Yaskawa INFORM job: THAPPY.JBI

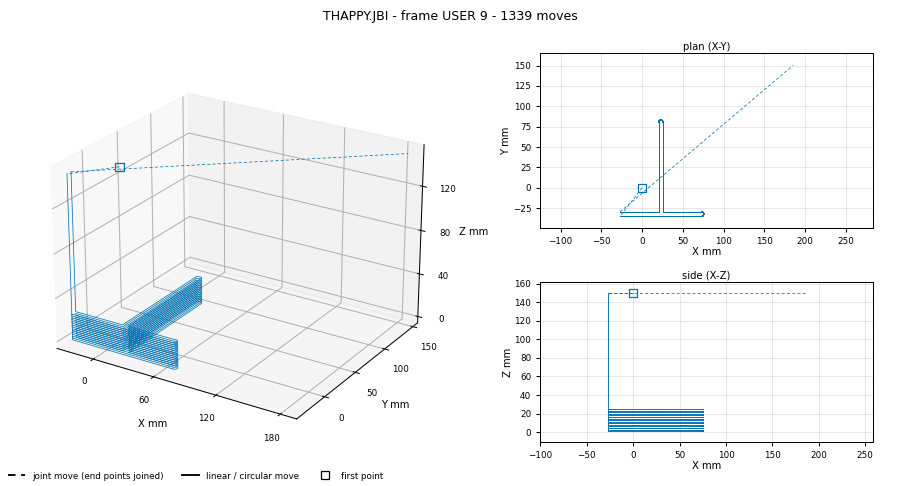
[picture p0: tool path of THAPPY.JBI in frame USER 9, 1339 of 1369 moves have a stored position in this frame; points joined in program order, loops and branches not executed]
/JOB
//NAME TTEST
//POS
///NPOS 1369,0,0,0,0,0
///USER 9
///TOOL 1
///POSTYPE USER
///RECTAN
///RCONF 1,0,0,0,0,0,0,0,0,0,0,0,0,0,0,0,0,0,0,0,0,0,0,0
C00000=0.000,0.000,150.000,0.0000,0.0000,-170.0000
C00001=-27.000,-35.000,150.000,0.0000,0.0000,-170.0000
C00002=-27.000,-35.000,1.000,0.0000,0.0000,-170.0000
C00003=-22.000,-35.000,1.000,0.0000,0.0000,-170.0000
C00004=-17.000,-35.000,1.000,0.0000,0.0000,-170.0000
C00005=-12.000,-35.000,1.000,0.0000,0.0000,-170.0000
C00006=-7.000,-35.000,1.000,0.0000,0.0000,-170.0000
C00007=-2.000,-35.000,1.000,0.0000,0.0000,-170.0000
C00008=3.000,-35.000,1.000,0.0000,0.0000,-170.0000
C00009=8.000,-35.000,1.000,0.0000,0.0000,-170.0000
C00010=13.000,-35.000,1.000,0.0000,0.0000,-170.0000
C00011=18.000,-35.000,1.000,0.0000,0.0000,-170.0000
C00012=23.000,-35.000,1.000,0.0000,0.0000,-170.0000
C00013=28.000,-35.000,1.000,0.0000,0.0000,-170.0000
C00014=33.000,-35.000,1.000,0.0000,0.0000,-170.0000
C00015=38.000,-35.000,1.000,0.0000,0.0000,-170.0000
C00016=43.000,-35.000,1.000,0.0000,0.0000,-170.0000
C00017=48.000,-35.000,1.000,0.0000,0.0000,-170.0000
C00018=53.000,-35.000,1.000,0.0000,0.0000,-170.0000
C00019=58.000,-35.000,1.000,0.0000,0.0000,-170.0000
C00020=63.000,-35.000,1.000,0.0000,0.0000,-170.0000
C00021=68.000,-35.000,1.000,0.0000,0.0000,-170.0000
C00022=73.000,-35.000,1.000,0.0000,0.0000,-170.0000
C00023=73.000,-35.000,1.000,0.0000,0.0000,-170.0000
C00024=75.750,-32.250,1.000,0.0000,0.0000,-170.0000
C00025=73.000,-29.500,1.000,0.0000,0.0000,-170.0000
C00026=68.275,-29.500,1.000,0.0000,0.0000,-170.0000
C00027=63.550,-29.500,1.000,0.0000,0.0000,-170.0000
C00028=58.825,-29.500,1.000,0.0000,0.0000,-170.0000
C00029=54.100,-29.500,1.000,0.0000,0.0000,-170.0000
C00030=49.375,-29.500,1.000,0.0000,0.0000,-170.0000
C00031=44.650,-29.500,1.000,0.0000,0.0000,-170.0000
C00032=39.925,-29.500,1.000,0.0000,0.0000,-170.0000
C00033=35.200,-29.500,1.000,0.0000,0.0000,-170.0000
C00034=30.475,-29.500,1.000,0.0000,0.0000,-170.0000
C00035=25.750,-29.500,1.000,0.0000,0.0000,-170.0000
C00036=25.750,-24.500,1.000,0.0000,0.0000,-170.0000
C00037=25.750,-19.500,1.000,0.0000,0.0000,-170.0000
C00038=25.750,-14.500,1.000,0.0000,0.0000,-170.0000
C00039=25.750,-9.500,1.000,0.0000,0.0000,-170.0000
C00040=25.750,-4.500,1.000,0.0000,0.0000,-170.0000
C00041=25.750,0.500,1.000,0.0000,0.0000,-170.0000
C00042=25.750,5.500,1.000,0.0000,0.0000,-170.0000
C00043=25.750,10.500,1.000,0.0000,0.0000,-170.0000
C00044=25.750,15.500,1.000,0.0000,0.0000,-170.0000
C00045=25.750,20.500,1.000,0.0000,0.0000,-170.0000
C00046=25.750,25.500,1.000,0.0000,0.0000,-170.0000
C00047=25.750,30.500,1.000,0.0000,0.0000,-170.0000
C00048=25.750,35.500,1.000,0.0000,0.0000,-170.0000
C00049=25.750,40.500,1.000,0.0000,0.0000,-170.0000
C00050=25.750,45.500,1.000,0.0000,0.0000,-170.0000
C00051=25.750,50.500,1.000,0.0000,0.0000,-170.0000
C00052=25.750,55.500,1.000,0.0000,0.0000,-170.0000
C00053=25.750,60.500,1.000,0.0000,0.0000,-170.0000
C00054=25.750,65.500,1.000,0.0000,0.0000,-170.0000
C00055=25.750,70.500,1.000,0.0000,0.0000,-170.0000
C00056=25.750,75.500,1.000,0.0000,0.0000,-170.0000
C00057=25.750,80.500,1.000,0.0000,0.0000,-170.0000
C00058=25.750,80.500,1.000,0.0000,0.0000,-170.0000
C00059=23.000,83.250,1.000,0.0000,0.0000,-170.0000
C00060=20.250,80.500,1.000,0.0000,0.0000,-170.0000
C00061=20.250,75.500,1.000,0.0000,0.0000,-170.0000
C00062=20.250,70.500,1.000,0.0000,0.0000,-170.0000
C00063=20.250,65.500,1.000,0.0000,0.0000,-170.0000
C00064=20.250,60.500,1.000,0.0000,0.0000,-170.0000
C00065=20.250,55.500,1.000,0.0000,0.0000,-170.0000
C00066=20.250,50.500,1.000,0.0000,0.0000,-170.0000
C00067=20.250,45.500,1.000,0.0000,0.0000,-170.0000
C00068=20.250,40.500,1.000,0.0000,0.0000,-170.0000
C00069=20.250,35.500,1.000,0.0000,0.0000,-170.0000
C00070=20.250,30.500,1.000,0.0000,0.0000,-170.0000
C00071=20.250,25.500,1.000,0.0000,0.0000,-170.0000
C00072=20.250,20.500,1.000,0.0000,0.0000,-170.0000
C00073=20.250,15.500,1.000,0.0000,0.0000,-170.0000
C00074=20.250,10.500,1.000,0.0000,0.0000,-170.0000
C00075=20.250,5.500,1.000,0.0000,0.0000,-170.0000
C00076=20.250,0.500,1.000,0.0000,0.0000,-170.0000
C00077=20.250,-4.500,1.000,0.0000,0.0000,-170.0000
C00078=20.250,-9.500,1.000,0.0000,0.0000,-170.0000
C00079=20.250,-14.500,1.000,0.0000,0.0000,-170.0000
C00080=20.250,-19.500,1.000,0.0000,0.0000,-170.0000
C00081=20.250,-24.500,1.000,0.0000,0.0000,-170.0000
C00082=20.250,-29.500,1.000,0.0000,0.0000,-170.0000
C00083=15.525,-29.500,1.000,0.0000,0.0000,-170.0000
C00084=10.800,-29.500,1.000,0.0000,0.0000,-170.0000
C00085=6.075,-29.500,1.000,0.0000,0.0000,-170.0000
C00086=1.350,-29.500,1.000,0.0000,0.0000,-170.0000
C00087=-3.375,-29.500,1.000,0.0000,0.0000,-170.0000
C00088=-8.100,-29.500,1.000,0.0000,0.0000,-170.0000
C00089=-12.825,-29.500,1.000,0.0000,0.0000,-170.0000
C00090=-17.550,-29.500,1.000,0.0000,0.0000,-170.0000
C00091=-22.275,-29.500,1.000,0.0000,0.0000,-170.0000
C00092=-27.000,-29.500,1.000,0.0000,0.0000,-170.0000
C00093=-27.000,-29.500,2.700,0.0000,0.0000,-170.0000
C00094=-22.275,-29.500,2.700,0.0000,0.0000,-170.0000
C00095=-17.550,-29.500,2.700,0.0000,0.0000,-170.0000
C00096=-12.825,-29.500,2.700,0.0000,0.0000,-170.0000
C00097=-8.100,-29.500,2.700,0.0000,0.0000,-170.0000
C00098=-3.375,-29.500,2.700,0.0000,0.0000,-170.0000
C00099=1.350,-29.500,2.700,0.0000,0.0000,-170.0000
C00100=6.075,-29.500,2.700,0.0000,0.0000,-170.0000
C00101=10.800,-29.500,2.700,0.0000,0.0000,-170.0000
C00102=15.525,-29.500,2.700,0.0000,0.0000,-170.0000
C00103=20.250,-29.500,2.700,0.0000,0.0000,-170.0000
C00104=20.250,-24.500,2.700,0.0000,0.0000,-170.0000
C00105=20.250,-19.500,2.700,0.0000,0.0000,-170.0000
C00106=20.250,-14.500,2.700,0.0000,0.0000,-170.0000
C00107=20.250,-9.500,2.700,0.0000,0.0000,-170.0000
C00108=20.250,-4.500,2.700,0.0000,0.0000,-170.0000
C00109=20.250,0.500,2.700,0.0000,0.0000,-170.0000
C00110=20.250,5.500,2.700,0.0000,0.0000,-170.0000
C00111=20.250,10.500,2.700,0.0000,0.0000,-170.0000
C00112=20.250,15.500,2.700,0.0000,0.0000,-170.0000
C00113=20.250,20.500,2.700,0.0000,0.0000,-170.0000
C00114=20.250,25.500,2.700,0.0000,0.0000,-170.0000
C00115=20.250,30.500,2.700,0.0000,0.0000,-170.0000
C00116=20.250,35.500,2.700,0.0000,0.0000,-170.0000
C00117=20.250,40.500,2.700,0.0000,0.0000,-170.0000
C00118=20.250,45.500,2.700,0.0000,0.0000,-170.0000
C00119=20.250,50.500,2.700,0.0000,0.0000,-170.0000
C00120=20.250,55.500,2.700,0.0000,0.0000,-170.0000
C00121=20.250,60.500,2.700,0.0000,0.0000,-170.0000
C00122=20.250,65.500,2.700,0.0000,0.0000,-170.0000
C00123=20.250,70.500,2.700,0.0000,0.0000,-170.0000
C00124=20.250,75.500,2.700,0.0000,0.0000,-170.0000
C00125=20.250,80.500,2.700,0.0000,0.0000,-170.0000
C00126=20.250,80.500,2.700,0.0000,0.0000,-170.0000
C00127=23.000,83.250,2.700,0.0000,0.0000,-170.0000
C00128=25.750,80.500,2.700,0.0000,0.0000,-170.0000
C00129=25.750,75.500,2.700,0.0000,0.0000,-170.0000
C00130=25.750,70.500,2.700,0.0000,0.0000,-170.0000
C00131=25.750,65.500,2.700,0.0000,0.0000,-170.0000
C00132=25.750,60.500,2.700,0.0000,0.0000,-170.0000
C00133=25.750,55.500,2.700,0.0000,0.0000,-170.0000
C00134=25.750,50.500,2.700,0.0000,0.0000,-170.0000
C00135=25.750,45.500,2.700,0.0000,0.0000,-170.0000
C00136=25.750,40.500,2.700,0.0000,0.0000,-170.0000
C00137=25.750,35.500,2.700,0.0000,0.0000,-170.0000
C00138=25.750,30.500,2.700,0.0000,0.0000,-170.0000
C00139=25.750,25.500,2.700,0.0000,0.0000,-170.0000
C00140=25.750,20.500,2.700,0.0000,0.0000,-170.0000
C00141=25.750,15.500,2.700,0.0000,0.0000,-170.0000
C00142=25.750,10.500,2.700,0.0000,0.0000,-170.0000
C00143=25.750,5.500,2.700,0.0000,0.0000,-170.0000
C00144=25.750,0.500,2.700,0.0000,0.0000,-170.0000
C00145=25.750,-4.500,2.700,0.0000,0.0000,-170.0000
C00146=25.750,-9.500,2.700,0.0000,0.0000,-170.0000
C00147=25.750,-14.500,2.700,0.0000,0.0000,-170.0000
C00148=25.750,-19.500,2.700,0.0000,0.0000,-170.0000
C00149=25.750,-24.500,2.700,0.0000,0.0000,-170.0000
C00150=25.750,-29.500,2.700,0.0000,0.0000,-170.0000
C00151=30.475,-29.500,2.700,0.0000,0.0000,-170.0000
C00152=35.200,-29.500,2.700,0.0000,0.0000,-170.0000
C00153=39.925,-29.500,2.700,0.0000,0.0000,-170.0000
C00154=44.650,-29.500,2.700,0.0000,0.0000,-170.0000
C00155=49.375,-29.500,2.700,0.0000,0.0000,-170.0000
C00156=54.100,-29.500,2.700,0.0000,0.0000,-170.0000
C00157=58.825,-29.500,2.700,0.0000,0.0000,-170.0000
C00158=63.550,-29.500,2.700,0.0000,0.0000,-170.0000
C00159=68.275,-29.500,2.700,0.0000,0.0000,-170.0000
C00160=73.000,-29.500,2.700,0.0000,0.0000,-170.0000
C00161=73.000,-29.500,2.700,0.0000,0.0000,-170.0000
C00162=75.750,-32.250,2.700,0.0000,0.0000,-170.0000
C00163=73.000,-35.000,2.700,0.0000,0.0000,-170.0000
C00164=68.000,-35.000,2.700,0.0000,0.0000,-170.0000
C00165=63.000,-35.000,2.700,0.0000,0.0000,-170.0000
C00166=58.000,-35.000,2.700,0.0000,0.0000,-170.0000
C00167=53.000,-35.000,2.700,0.0000,0.0000,-170.0000
C00168=48.000,-35.000,2.700,0.0000,0.0000,-170.0000
C00169=43.000,-35.000,2.700,0.0000,0.0000,-170.0000
C00170=38.000,-35.000,2.700,0.0000,0.0000,-170.0000
C00171=33.000,-35.000,2.700,0.0000,0.0000,-170.0000
C00172=28.000,-35.000,2.700,0.0000,0.0000,-170.0000
C00173=23.000,-35.000,2.700,0.0000,0.0000,-170.0000
C00174=18.000,-35.000,2.700,0.0000,0.0000,-170.0000
C00175=13.000,-35.000,2.700,0.0000,0.0000,-170.0000
C00176=8.000,-35.000,2.700,0.0000,0.0000,-170.0000
C00177=3.000,-35.000,2.700,0.0000,0.0000,-170.0000
C00178=-2.000,-35.000,2.700,0.0000,0.0000,-170.0000
C00179=-7.000,-35.000,2.700,0.0000,0.0000,-170.0000
C00180=-12.000,-35.000,2.700,0.0000,0.0000,-170.0000
C00181=-17.000,-35.000,2.700,0.0000,0.0000,-170.0000
C00182=-22.000,-35.000,2.700,0.0000,0.0000,-170.0000
C00183=-27.000,-35.000,2.700,0.0000,0.0000,-170.0000
C00184=-27.000,-35.000,4.400,0.0000,0.0000,-170.0000
C00185=-22.000,-35.000,4.400,0.0000,0.0000,-170.0000
C00186=-17.000,-35.000,4.400,0.0000,0.0000,-170.0000
C00187=-12.000,-35.000,4.400,0.0000,0.0000,-170.0000
C00188=-7.000,-35.000,4.400,0.0000,0.0000,-170.0000
C00189=-2.000,-35.000,4.400,0.0000,0.0000,-170.0000
C00190=3.000,-35.000,4.400,0.0000,0.0000,-170.0000
C00191=8.000,-35.000,4.400,0.0000,0.0000,-170.0000
C00192=13.000,-35.000,4.400,0.0000,0.0000,-170.0000
C00193=18.000,-35.000,4.400,0.0000,0.0000,-170.0000
C00194=23.000,-35.000,4.400,0.0000,0.0000,-170.0000
C00195=28.000,-35.000,4.400,0.0000,0.0000,-170.0000
C00196=33.000,-35.000,4.400,0.0000,0.0000,-170.0000
C00197=38.000,-35.000,4.400,0.0000,0.0000,-170.0000
C00198=43.000,-35.000,4.400,0.0000,0.0000,-170.0000
C00199=48.000,-35.000,4.400,0.0000,0.0000,-170.0000
C00200=53.000,-35.000,4.400,0.0000,0.0000,-170.0000
C00201=58.000,-35.000,4.400,0.0000,0.0000,-170.0000
C00202=63.000,-35.000,4.400,0.0000,0.0000,-170.0000
C00203=68.000,-35.000,4.400,0.0000,0.0000,-170.0000
C00204=73.000,-35.000,4.400,0.0000,0.0000,-170.0000
C00205=73.000,-35.000,4.400,0.0000,0.0000,-170.0000
C00206=75.750,-32.250,4.400,0.0000,0.0000,-170.0000
C00207=73.000,-29.500,4.400,0.0000,0.0000,-170.0000
C00208=68.275,-29.500,4.400,0.0000,0.0000,-170.0000
C00209=63.550,-29.500,4.400,0.0000,0.0000,-170.0000
C00210=58.825,-29.500,4.400,0.0000,0.0000,-170.0000
C00211=54.100,-29.500,4.400,0.0000,0.0000,-170.0000
C00212=49.375,-29.500,4.400,0.0000,0.0000,-170.0000
C00213=44.650,-29.500,4.400,0.0000,0.0000,-170.0000
C00214=39.925,-29.500,4.400,0.0000,0.0000,-170.0000
C00215=35.200,-29.500,4.400,0.0000,0.0000,-170.0000
C00216=30.475,-29.500,4.400,0.0000,0.0000,-170.0000
C00217=25.750,-29.500,4.400,0.0000,0.0000,-170.0000
C00218=25.750,-24.500,4.400,0.0000,0.0000,-170.0000
C00219=25.750,-19.500,4.400,0.0000,0.0000,-170.0000
C00220=25.750,-14.500,4.400,0.0000,0.0000,-170.0000
C00221=25.750,-9.500,4.400,0.0000,0.0000,-170.0000
C00222=25.750,-4.500,4.400,0.0000,0.0000,-170.0000
C00223=25.750,0.500,4.400,0.0000,0.0000,-170.0000
C00224=25.750,5.500,4.400,0.0000,0.0000,-170.0000
C00225=25.750,10.500,4.400,0.0000,0.0000,-170.0000
C00226=25.750,15.500,4.400,0.0000,0.0000,-170.0000
C00227=25.750,20.500,4.400,0.0000,0.0000,-170.0000
C00228=25.750,25.500,4.400,0.0000,0.0000,-170.0000
C00229=25.750,30.500,4.400,0.0000,0.0000,-170.0000
C00230=25.750,35.500,4.400,0.0000,0.0000,-170.0000
C00231=25.750,40.500,4.400,0.0000,0.0000,-170.0000
C00232=25.750,45.500,4.400,0.0000,0.0000,-170.0000
C00233=25.750,50.500,4.400,0.0000,0.0000,-170.0000
C00234=25.750,55.500,4.400,0.0000,0.0000,-170.0000
C00235=25.750,60.500,4.400,0.0000,0.0000,-170.0000
C00236=25.750,65.500,4.400,0.0000,0.0000,-170.0000
C00237=25.750,70.500,4.400,0.0000,0.0000,-170.0000
C00238=25.750,75.500,4.400,0.0000,0.0000,-170.0000
C00239=25.750,80.500,4.400,0.0000,0.0000,-170.0000
C00240=25.750,80.500,4.400,0.0000,0.0000,-170.0000
C00241=23.000,83.250,4.400,0.0000,0.0000,-170.0000
C00242=20.250,80.500,4.400,0.0000,0.0000,-170.0000
C00243=20.250,75.500,4.400,0.0000,0.0000,-170.0000
C00244=20.250,70.500,4.400,0.0000,0.0000,-170.0000
C00245=20.250,65.500,4.400,0.0000,0.0000,-170.0000
C00246=20.250,60.500,4.400,0.0000,0.0000,-170.0000
C00247=20.250,55.500,4.400,0.0000,0.0000,-170.0000
C00248=20.250,50.500,4.400,0.0000,0.0000,-170.0000
C00249=20.250,45.500,4.400,0.0000,0.0000,-170.0000
C00250=20.250,40.500,4.400,0.0000,0.0000,-170.0000
C00251=20.250,35.500,4.400,0.0000,0.0000,-170.0000
C00252=20.250,30.500,4.400,0.0000,0.0000,-170.0000
C00253=20.250,25.500,4.400,0.0000,0.0000,-170.0000
C00254=20.250,20.500,4.400,0.0000,0.0000,-170.0000
C00255=20.250,15.500,4.400,0.0000,0.0000,-170.0000
C00256=20.250,10.500,4.400,0.0000,0.0000,-170.0000
C00257=20.250,5.500,4.400,0.0000,0.0000,-170.0000
C00258=20.250,0.500,4.400,0.0000,0.0000,-170.0000
C00259=20.250,-4.500,4.400,0.0000,0.0000,-170.0000
C00260=20.250,-9.500,4.400,0.0000,0.0000,-170.0000
C00261=20.250,-14.500,4.400,0.0000,0.0000,-170.0000
C00262=20.250,-19.500,4.400,0.0000,0.0000,-170.0000
C00263=20.250,-24.500,4.400,0.0000,0.0000,-170.0000
C00264=20.250,-29.500,4.400,0.0000,0.0000,-170.0000
C00265=15.525,-29.500,4.400,0.0000,0.0000,-170.0000
C00266=10.800,-29.500,4.400,0.0000,0.0000,-170.0000
C00267=6.075,-29.500,4.400,0.0000,0.0000,-170.0000
C00268=1.350,-29.500,4.400,0.0000,0.0000,-170.0000
C00269=-3.375,-29.500,4.400,0.0000,0.0000,-170.0000
C00270=-8.100,-29.500,4.400,0.0000,0.0000,-170.0000
C00271=-12.825,-29.500,4.400,0.0000,0.0000,-170.0000
C00272=-17.550,-29.500,4.400,0.0000,0.0000,-170.0000
C00273=-22.275,-29.500,4.400,0.0000,0.0000,-170.0000
C00274=-27.000,-29.500,4.400,0.0000,0.0000,-170.0000
C00275=-27.000,-29.500,6.100,0.0000,0.0000,-170.0000
C00276=-22.275,-29.500,6.100,0.0000,0.0000,-170.0000
C00277=-17.550,-29.500,6.100,0.0000,0.0000,-170.0000
C00278=-12.825,-29.500,6.100,0.0000,0.0000,-170.0000
C00279=-8.100,-29.500,6.100,0.0000,0.0000,-170.0000
C00280=-3.375,-29.500,6.100,0.0000,0.0000,-170.0000
C00281=1.350,-29.500,6.100,0.0000,0.0000,-170.0000
C00282=6.075,-29.500,6.100,0.0000,0.0000,-170.0000
C00283=10.800,-29.500,6.100,0.0000,0.0000,-170.0000
C00284=15.525,-29.500,6.100,0.0000,0.0000,-170.0000
C00285=20.250,-29.500,6.100,0.0000,0.0000,-170.0000
C00286=20.250,-24.500,6.100,0.0000,0.0000,-170.0000
C00287=20.250,-19.500,6.100,0.0000,0.0000,-170.0000
C00288=20.250,-14.500,6.100,0.0000,0.0000,-170.0000
C00289=20.250,-9.500,6.100,0.0000,0.0000,-170.0000
C00290=20.250,-4.500,6.100,0.0000,0.0000,-170.0000
C00291=20.250,0.500,6.100,0.0000,0.0000,-170.0000
C00292=20.250,5.500,6.100,0.0000,0.0000,-170.0000
C00293=20.250,10.500,6.100,0.0000,0.0000,-170.0000
C00294=20.250,15.500,6.100,0.0000,0.0000,-170.0000
C00295=20.250,20.500,6.100,0.0000,0.0000,-170.0000
C00296=20.250,25.500,6.100,0.0000,0.0000,-170.0000
C00297=20.250,30.500,6.100,0.0000,0.0000,-170.0000
C00298=20.250,35.500,6.100,0.0000,0.0000,-170.0000
C00299=20.250,40.500,6.100,0.0000,0.0000,-170.0000
C00300=20.250,45.500,6.100,0.0000,0.0000,-170.0000
C00301=20.250,50.500,6.100,0.0000,0.0000,-170.0000
C00302=20.250,55.500,6.100,0.0000,0.0000,-170.0000
C00303=20.250,60.500,6.100,0.0000,0.0000,-170.0000
C00304=20.250,65.500,6.100,0.0000,0.0000,-170.0000
C00305=20.250,70.500,6.100,0.0000,0.0000,-170.0000
C00306=20.250,75.500,6.100,0.0000,0.0000,-170.0000
C00307=20.250,80.500,6.100,0.0000,0.0000,-170.0000
C00308=20.250,80.500,6.100,0.0000,0.0000,-170.0000
C00309=23.000,83.250,6.100,0.0000,0.0000,-170.0000
C00310=25.750,80.500,6.100,0.0000,0.0000,-170.0000
C00311=25.750,75.500,6.100,0.0000,0.0000,-170.0000
C00312=25.750,70.500,6.100,0.0000,0.0000,-170.0000
C00313=25.750,65.500,6.100,0.0000,0.0000,-170.0000
C00314=25.750,60.500,6.100,0.0000,0.0000,-170.0000
C00315=25.750,55.500,6.100,0.0000,0.0000,-170.0000
C00316=25.750,50.500,6.100,0.0000,0.0000,-170.0000
C00317=25.750,45.500,6.100,0.0000,0.0000,-170.0000
C00318=25.750,40.500,6.100,0.0000,0.0000,-170.0000
C00319=25.750,35.500,6.100,0.0000,0.0000,-170.0000
C00320=25.750,30.500,6.100,0.0000,0.0000,-170.0000
C00321=25.750,25.500,6.100,0.0000,0.0000,-170.0000
C00322=25.750,20.500,6.100,0.0000,0.0000,-170.0000
C00323=25.750,15.500,6.100,0.0000,0.0000,-170.0000
C00324=25.750,10.500,6.100,0.0000,0.0000,-170.0000
C00325=25.750,5.500,6.100,0.0000,0.0000,-170.0000
C00326=25.750,0.500,6.100,0.0000,0.0000,-170.0000
C00327=25.750,-4.500,6.100,0.0000,0.0000,-170.0000
C00328=25.750,-9.500,6.100,0.0000,0.0000,-170.0000
C00329=25.750,-14.500,6.100,0.0000,0.0000,-170.0000
C00330=25.750,-19.500,6.100,0.0000,0.0000,-170.0000
C00331=25.750,-24.500,6.100,0.0000,0.0000,-170.0000
C00332=25.750,-29.500,6.100,0.0000,0.0000,-170.0000
C00333=30.475,-29.500,6.100,0.0000,0.0000,-170.0000
C00334=35.200,-29.500,6.100,0.0000,0.0000,-170.0000
C00335=39.925,-29.500,6.100,0.0000,0.0000,-170.0000
C00336=44.650,-29.500,6.100,0.0000,0.0000,-170.0000
C00337=49.375,-29.500,6.100,0.0000,0.0000,-170.0000
C00338=54.100,-29.500,6.100,0.0000,0.0000,-170.0000
C00339=58.825,-29.500,6.100,0.0000,0.0000,-170.0000
C00340=63.550,-29.500,6.100,0.0000,0.0000,-170.0000
C00341=68.275,-29.500,6.100,0.0000,0.0000,-170.0000
C00342=73.000,-29.500,6.100,0.0000,0.0000,-170.0000
C00343=73.000,-29.500,6.100,0.0000,0.0000,-170.0000
C00344=75.750,-32.250,6.100,0.0000,0.0000,-170.0000
C00345=73.000,-35.000,6.100,0.0000,0.0000,-170.0000
C00346=68.000,-35.000,6.100,0.0000,0.0000,-170.0000
C00347=63.000,-35.000,6.100,0.0000,0.0000,-170.0000
C00348=58.000,-35.000,6.100,0.0000,0.0000,-170.0000
C00349=53.000,-35.000,6.100,0.0000,0.0000,-170.0000
C00350=48.000,-35.000,6.100,0.0000,0.0000,-170.0000
C00351=43.000,-35.000,6.100,0.0000,0.0000,-170.0000
C00352=38.000,-35.000,6.100,0.0000,0.0000,-170.0000
C00353=33.000,-35.000,6.100,0.0000,0.0000,-170.0000
C00354=28.000,-35.000,6.100,0.0000,0.0000,-170.0000
C00355=23.000,-35.000,6.100,0.0000,0.0000,-170.0000
C00356=18.000,-35.000,6.100,0.0000,0.0000,-170.0000
C00357=13.000,-35.000,6.100,0.0000,0.0000,-170.0000
C00358=8.000,-35.000,6.100,0.0000,0.0000,-170.0000
C00359=3.000,-35.000,6.100,0.0000,0.0000,-170.0000
C00360=-2.000,-35.000,6.100,0.0000,0.0000,-170.0000
C00361=-7.000,-35.000,6.100,0.0000,0.0000,-170.0000
C00362=-12.000,-35.000,6.100,0.0000,0.0000,-170.0000
C00363=-17.000,-35.000,6.100,0.0000,0.0000,-170.0000
C00364=-22.000,-35.000,6.100,0.0000,0.0000,-170.0000
C00365=-27.000,-35.000,6.100,0.0000,0.0000,-170.0000
C00366=-27.000,-35.000,7.800,0.0000,0.0000,-170.0000
C00367=-22.000,-35.000,7.800,0.0000,0.0000,-170.0000
C00368=-17.000,-35.000,7.800,0.0000,0.0000,-170.0000
C00369=-12.000,-35.000,7.800,0.0000,0.0000,-170.0000
C00370=-7.000,-35.000,7.800,0.0000,0.0000,-170.0000
C00371=-2.000,-35.000,7.800,0.0000,0.0000,-170.0000
C00372=3.000,-35.000,7.800,0.0000,0.0000,-170.0000
C00373=8.000,-35.000,7.800,0.0000,0.0000,-170.0000
C00374=13.000,-35.000,7.800,0.0000,0.0000,-170.0000
C00375=18.000,-35.000,7.800,0.0000,0.0000,-170.0000
C00376=23.000,-35.000,7.800,0.0000,0.0000,-170.0000
C00377=28.000,-35.000,7.800,0.0000,0.0000,-170.0000
C00378=33.000,-35.000,7.800,0.0000,0.0000,-170.0000
C00379=38.000,-35.000,7.800,0.0000,0.0000,-170.0000
C00380=43.000,-35.000,7.800,0.0000,0.0000,-170.0000
C00381=48.000,-35.000,7.800,0.0000,0.0000,-170.0000
C00382=53.000,-35.000,7.800,0.0000,0.0000,-170.0000
C00383=58.000,-35.000,7.800,0.0000,0.0000,-170.0000
C00384=63.000,-35.000,7.800,0.0000,0.0000,-170.0000
C00385=68.000,-35.000,7.800,0.0000,0.0000,-170.0000
C00386=73.000,-35.000,7.800,0.0000,0.0000,-170.0000
C00387=73.000,-35.000,7.800,0.0000,0.0000,-170.0000
C00388=75.750,-32.250,7.800,0.0000,0.0000,-170.0000
C00389=73.000,-29.500,7.800,0.0000,0.0000,-170.0000
C00390=68.275,-29.500,7.800,0.0000,0.0000,-170.0000
C00391=63.550,-29.500,7.800,0.0000,0.0000,-170.0000
C00392=58.825,-29.500,7.800,0.0000,0.0000,-170.0000
C00393=54.100,-29.500,7.800,0.0000,0.0000,-170.0000
C00394=49.375,-29.500,7.800,0.0000,0.0000,-170.0000
C00395=44.650,-29.500,7.800,0.0000,0.0000,-170.0000
C00396=39.925,-29.500,7.800,0.0000,0.0000,-170.0000
C00397=35.200,-29.500,7.800,0.0000,0.0000,-170.0000
C00398=30.475,-29.500,7.800,0.0000,0.0000,-170.0000
C00399=25.750,-29.500,7.800,0.0000,0.0000,-170.0000
C00400=25.750,-24.500,7.800,0.0000,0.0000,-170.0000
C00401=25.750,-19.500,7.800,0.0000,0.0000,-170.0000
C00402=25.750,-14.500,7.800,0.0000,0.0000,-170.0000
C00403=25.750,-9.500,7.800,0.0000,0.0000,-170.0000
C00404=25.750,-4.500,7.800,0.0000,0.0000,-170.0000
C00405=25.750,0.500,7.800,0.0000,0.0000,-170.0000
C00406=25.750,5.500,7.800,0.0000,0.0000,-170.0000
C00407=25.750,10.500,7.800,0.0000,0.0000,-170.0000
C00408=25.750,15.500,7.800,0.0000,0.0000,-170.0000
C00409=25.750,20.500,7.800,0.0000,0.0000,-170.0000
C00410=25.750,25.500,7.800,0.0000,0.0000,-170.0000
C00411=25.750,30.500,7.800,0.0000,0.0000,-170.0000
C00412=25.750,35.500,7.800,0.0000,0.0000,-170.0000
C00413=25.750,40.500,7.800,0.0000,0.0000,-170.0000
C00414=25.750,45.500,7.800,0.0000,0.0000,-170.0000
C00415=25.750,50.500,7.800,0.0000,0.0000,-170.0000
C00416=25.750,55.500,7.800,0.0000,0.0000,-170.0000
C00417=25.750,60.500,7.800,0.0000,0.0000,-170.0000
C00418=25.750,65.500,7.800,0.0000,0.0000,-170.0000
C00419=25.750,70.500,7.800,0.0000,0.0000,-170.0000
C00420=25.750,75.500,7.800,0.0000,0.0000,-170.0000
C00421=25.750,80.500,7.800,0.0000,0.0000,-170.0000
C00422=25.750,80.500,7.800,0.0000,0.0000,-170.0000
C00423=23.000,83.250,7.800,0.0000,0.0000,-170.0000
C00424=20.250,80.500,7.800,0.0000,0.0000,-170.0000
C00425=20.250,75.500,7.800,0.0000,0.0000,-170.0000
C00426=20.250,70.500,7.800,0.0000,0.0000,-170.0000
C00427=20.250,65.500,7.800,0.0000,0.0000,-170.0000
C00428=20.250,60.500,7.800,0.0000,0.0000,-170.0000
C00429=20.250,55.500,7.800,0.0000,0.0000,-170.0000
C00430=20.250,50.500,7.800,0.0000,0.0000,-170.0000
C00431=20.250,45.500,7.800,0.0000,0.0000,-170.0000
C00432=20.250,40.500,7.800,0.0000,0.0000,-170.0000
C00433=20.250,35.500,7.800,0.0000,0.0000,-170.0000
C00434=20.250,30.500,7.800,0.0000,0.0000,-170.0000
C00435=20.250,25.500,7.800,0.0000,0.0000,-170.0000
C00436=20.250,20.500,7.800,0.0000,0.0000,-170.0000
C00437=20.250,15.500,7.800,0.0000,0.0000,-170.0000
C00438=20.250,10.500,7.800,0.0000,0.0000,-170.0000
C00439=20.250,5.500,7.800,0.0000,0.0000,-170.0000
C00440=20.250,0.500,7.800,0.0000,0.0000,-170.0000
C00441=20.250,-4.500,7.800,0.0000,0.0000,-170.0000
C00442=20.250,-9.500,7.800,0.0000,0.0000,-170.0000
C00443=20.250,-14.500,7.800,0.0000,0.0000,-170.0000
C00444=20.250,-19.500,7.800,0.0000,0.0000,-170.0000
C00445=20.250,-24.500,7.800,0.0000,0.0000,-170.0000
C00446=20.250,-29.500,7.800,0.0000,0.0000,-170.0000
C00447=15.525,-29.500,7.800,0.0000,0.0000,-170.0000
C00448=10.800,-29.500,7.800,0.0000,0.0000,-170.0000
C00449=6.075,-29.500,7.800,0.0000,0.0000,-170.0000
C00450=1.350,-29.500,7.800,0.0000,0.0000,-170.0000
C00451=-3.375,-29.500,7.800,0.0000,0.0000,-170.0000
C00452=-8.100,-29.500,7.800,0.0000,0.0000,-170.0000
C00453=-12.825,-29.500,7.800,0.0000,0.0000,-170.0000
C00454=-17.550,-29.500,7.800,0.0000,0.0000,-170.0000
C00455=-22.275,-29.500,7.800,0.0000,0.0000,-170.0000
C00456=-27.000,-29.500,7.800,0.0000,0.0000,-170.0000
C00457=-27.000,-29.500,9.500,0.0000,0.0000,-170.0000
C00458=-22.275,-29.500,9.500,0.0000,0.0000,-170.0000
C00459=-17.550,-29.500,9.500,0.0000,0.0000,-170.0000
C00460=-12.825,-29.500,9.500,0.0000,0.0000,-170.0000
C00461=-8.100,-29.500,9.500,0.0000,0.0000,-170.0000
C00462=-3.375,-29.500,9.500,0.0000,0.0000,-170.0000
C00463=1.350,-29.500,9.500,0.0000,0.0000,-170.0000
C00464=6.075,-29.500,9.500,0.0000,0.0000,-170.0000
C00465=10.800,-29.500,9.500,0.0000,0.0000,-170.0000
C00466=15.525,-29.500,9.500,0.0000,0.0000,-170.0000
C00467=20.250,-29.500,9.500,0.0000,0.0000,-170.0000
C00468=20.250,-24.500,9.500,0.0000,0.0000,-170.0000
C00469=20.250,-19.500,9.500,0.0000,0.0000,-170.0000
C00470=20.250,-14.500,9.500,0.0000,0.0000,-170.0000
C00471=20.250,-9.500,9.500,0.0000,0.0000,-170.0000
C00472=20.250,-4.500,9.500,0.0000,0.0000,-170.0000
C00473=20.250,0.500,9.500,0.0000,0.0000,-170.0000
C00474=20.250,5.500,9.500,0.0000,0.0000,-170.0000
C00475=20.250,10.500,9.500,0.0000,0.0000,-170.0000
C00476=20.250,15.500,9.500,0.0000,0.0000,-170.0000
C00477=20.250,20.500,9.500,0.0000,0.0000,-170.0000
C00478=20.250,25.500,9.500,0.0000,0.0000,-170.0000
C00479=20.250,30.500,9.500,0.0000,0.0000,-170.0000
C00480=20.250,35.500,9.500,0.0000,0.0000,-170.0000
C00481=20.250,40.500,9.500,0.0000,0.0000,-170.0000
C00482=20.250,45.500,9.500,0.0000,0.0000,-170.0000
C00483=20.250,50.500,9.500,0.0000,0.0000,-170.0000
C00484=20.250,55.500,9.500,0.0000,0.0000,-170.0000
C00485=20.250,60.500,9.500,0.0000,0.0000,-170.0000
C00486=20.250,65.500,9.500,0.0000,0.0000,-170.0000
C00487=20.250,70.500,9.500,0.0000,0.0000,-170.0000
C00488=20.250,75.500,9.500,0.0000,0.0000,-170.0000
C00489=20.250,80.500,9.500,0.0000,0.0000,-170.0000
C00490=20.250,80.500,9.500,0.0000,0.0000,-170.0000
C00491=23.000,83.250,9.500,0.0000,0.0000,-170.0000
C00492=25.750,80.500,9.500,0.0000,0.0000,-170.0000
C00493=25.750,75.500,9.500,0.0000,0.0000,-170.0000
C00494=25.750,70.500,9.500,0.0000,0.0000,-170.0000
C00495=25.750,65.500,9.500,0.0000,0.0000,-170.0000
C00496=25.750,60.500,9.500,0.0000,0.0000,-170.0000
C00497=25.750,55.500,9.500,0.0000,0.0000,-170.0000
C00498=25.750,50.500,9.500,0.0000,0.0000,-170.0000
C00499=25.750,45.500,9.500,0.0000,0.0000,-170.0000
C00500=25.750,40.500,9.500,0.0000,0.0000,-170.0000
C00501=25.750,35.500,9.500,0.0000,0.0000,-170.0000
C00502=25.750,30.500,9.500,0.0000,0.0000,-170.0000
C00503=25.750,25.500,9.500,0.0000,0.0000,-170.0000
C00504=25.750,20.500,9.500,0.0000,0.0000,-170.0000
C00505=25.750,15.500,9.500,0.0000,0.0000,-170.0000
C00506=25.750,10.500,9.500,0.0000,0.0000,-170.0000
C00507=25.750,5.500,9.500,0.0000,0.0000,-170.0000
C00508=25.750,0.500,9.500,0.0000,0.0000,-170.0000
C00509=25.750,-4.500,9.500,0.0000,0.0000,-170.0000
C00510=25.750,-9.500,9.500,0.0000,0.0000,-170.0000
C00511=25.750,-14.500,9.500,0.0000,0.0000,-170.0000
C00512=25.750,-19.500,9.500,0.0000,0.0000,-170.0000
C00513=25.750,-24.500,9.500,0.0000,0.0000,-170.0000
C00514=25.750,-29.500,9.500,0.0000,0.0000,-170.0000
C00515=30.475,-29.500,9.500,0.0000,0.0000,-170.0000
C00516=35.200,-29.500,9.500,0.0000,0.0000,-170.0000
C00517=39.925,-29.500,9.500,0.0000,0.0000,-170.0000
C00518=44.650,-29.500,9.500,0.0000,0.0000,-170.0000
C00519=49.375,-29.500,9.500,0.0000,0.0000,-170.0000
C00520=54.100,-29.500,9.500,0.0000,0.0000,-170.0000
C00521=58.825,-29.500,9.500,0.0000,0.0000,-170.0000
C00522=63.550,-29.500,9.500,0.0000,0.0000,-170.0000
C00523=68.275,-29.500,9.500,0.0000,0.0000,-170.0000
C00524=73.000,-29.500,9.500,0.0000,0.0000,-170.0000
C00525=73.000,-29.500,9.500,0.0000,0.0000,-170.0000
C00526=75.750,-32.250,9.500,0.0000,0.0000,-170.0000
C00527=73.000,-35.000,9.500,0.0000,0.0000,-170.0000
C00528=68.000,-35.000,9.500,0.0000,0.0000,-170.0000
C00529=63.000,-35.000,9.500,0.0000,0.0000,-170.0000
C00530=58.000,-35.000,9.500,0.0000,0.0000,-170.0000
C00531=53.000,-35.000,9.500,0.0000,0.0000,-170.0000
C00532=48.000,-35.000,9.500,0.0000,0.0000,-170.0000
C00533=43.000,-35.000,9.500,0.0000,0.0000,-170.0000
C00534=38.000,-35.000,9.500,0.0000,0.0000,-170.0000
C00535=33.000,-35.000,9.500,0.0000,0.0000,-170.0000
C00536=28.000,-35.000,9.500,0.0000,0.0000,-170.0000
C00537=23.000,-35.000,9.500,0.0000,0.0000,-170.0000
C00538=18.000,-35.000,9.500,0.0000,0.0000,-170.0000
C00539=13.000,-35.000,9.500,0.0000,0.0000,-170.0000
C00540=8.000,-35.000,9.500,0.0000,0.0000,-170.0000
C00541=3.000,-35.000,9.500,0.0000,0.0000,-170.0000
C00542=-2.000,-35.000,9.500,0.0000,0.0000,-170.0000
C00543=-7.000,-35.000,9.500,0.0000,0.0000,-170.0000
C00544=-12.000,-35.000,9.500,0.0000,0.0000,-170.0000
C00545=-17.000,-35.000,9.500,0.0000,0.0000,-170.0000
C00546=-22.000,-35.000,9.500,0.0000,0.0000,-170.0000
C00547=-27.000,-35.000,9.500,0.0000,0.0000,-170.0000
C00548=-27.000,-35.000,11.200,0.0000,0.0000,-170.0000
C00549=-22.000,-35.000,11.200,0.0000,0.0000,-170.0000
C00550=-17.000,-35.000,11.200,0.0000,0.0000,-170.0000
C00551=-12.000,-35.000,11.200,0.0000,0.0000,-170.0000
C00552=-7.000,-35.000,11.200,0.0000,0.0000,-170.0000
C00553=-2.000,-35.000,11.200,0.0000,0.0000,-170.0000
C00554=3.000,-35.000,11.200,0.0000,0.0000,-170.0000
C00555=8.000,-35.000,11.200,0.0000,0.0000,-170.0000
C00556=13.000,-35.000,11.200,0.0000,0.0000,-170.0000
C00557=18.000,-35.000,11.200,0.0000,0.0000,-170.0000
C00558=23.000,-35.000,11.200,0.0000,0.0000,-170.0000
C00559=28.000,-35.000,11.200,0.0000,0.0000,-170.0000
C00560=33.000,-35.000,11.200,0.0000,0.0000,-170.0000
C00561=38.000,-35.000,11.200,0.0000,0.0000,-170.0000
C00562=43.000,-35.000,11.200,0.0000,0.0000,-170.0000
C00563=48.000,-35.000,11.200,0.0000,0.0000,-170.0000
C00564=53.000,-35.000,11.200,0.0000,0.0000,-170.0000
C00565=58.000,-35.000,11.200,0.0000,0.0000,-170.0000
C00566=63.000,-35.000,11.200,0.0000,0.0000,-170.0000
C00567=68.000,-35.000,11.200,0.0000,0.0000,-170.0000
C00568=73.000,-35.000,11.200,0.0000,0.0000,-170.0000
C00569=73.000,-35.000,11.200,0.0000,0.0000,-170.0000
C00570=75.750,-32.250,11.200,0.0000,0.0000,-170.0000
C00571=73.000,-29.500,11.200,0.0000,0.0000,-170.0000
C00572=68.275,-29.500,11.200,0.0000,0.0000,-170.0000
C00573=63.550,-29.500,11.200,0.0000,0.0000,-170.0000
C00574=58.825,-29.500,11.200,0.0000,0.0000,-170.0000
C00575=54.100,-29.500,11.200,0.0000,0.0000,-170.0000
C00576=49.375,-29.500,11.200,0.0000,0.0000,-170.0000
C00577=44.650,-29.500,11.200,0.0000,0.0000,-170.0000
C00578=39.925,-29.500,11.200,0.0000,0.0000,-170.0000
C00579=35.200,-29.500,11.200,0.0000,0.0000,-170.0000
C00580=30.475,-29.500,11.200,0.0000,0.0000,-170.0000
C00581=25.750,-29.500,11.200,0.0000,0.0000,-170.0000
C00582=25.750,-24.500,11.200,0.0000,0.0000,-170.0000
C00583=25.750,-19.500,11.200,0.0000,0.0000,-170.0000
C00584=25.750,-14.500,11.200,0.0000,0.0000,-170.0000
C00585=25.750,-9.500,11.200,0.0000,0.0000,-170.0000
C00586=25.750,-4.500,11.200,0.0000,0.0000,-170.0000
C00587=25.750,0.500,11.200,0.0000,0.0000,-170.0000
C00588=25.750,5.500,11.200,0.0000,0.0000,-170.0000
C00589=25.750,10.500,11.200,0.0000,0.0000,-170.0000
C00590=25.750,15.500,11.200,0.0000,0.0000,-170.0000
C00591=25.750,20.500,11.200,0.0000,0.0000,-170.0000
C00592=25.750,25.500,11.200,0.0000,0.0000,-170.0000
C00593=25.750,30.500,11.200,0.0000,0.0000,-170.0000
C00594=25.750,35.500,11.200,0.0000,0.0000,-170.0000
C00595=25.750,40.500,11.200,0.0000,0.0000,-170.0000
C00596=25.750,45.500,11.200,0.0000,0.0000,-170.0000
C00597=25.750,50.500,11.200,0.0000,0.0000,-170.0000
C00598=25.750,55.500,11.200,0.0000,0.0000,-170.0000
C00599=25.750,60.500,11.200,0.0000,0.0000,-170.0000
C00600=25.750,65.500,11.200,0.0000,0.0000,-170.0000
C00601=25.750,70.500,11.200,0.0000,0.0000,-170.0000
C00602=25.750,75.500,11.200,0.0000,0.0000,-170.0000
C00603=25.750,80.500,11.200,0.0000,0.0000,-170.0000
C00604=25.750,80.500,11.200,0.0000,0.0000,-170.0000
C00605=23.000,83.250,11.200,0.0000,0.0000,-170.0000
C00606=20.250,80.500,11.200,0.0000,0.0000,-170.0000
C00607=20.250,75.500,11.200,0.0000,0.0000,-170.0000
C00608=20.250,70.500,11.200,0.0000,0.0000,-170.0000
C00609=20.250,65.500,11.200,0.0000,0.0000,-170.0000
C00610=20.250,60.500,11.200,0.0000,0.0000,-170.0000
C00611=20.250,55.500,11.200,0.0000,0.0000,-170.0000
C00612=20.250,50.500,11.200,0.0000,0.0000,-170.0000
C00613=20.250,45.500,11.200,0.0000,0.0000,-170.0000
C00614=20.250,40.500,11.200,0.0000,0.0000,-170.0000
C00615=20.250,35.500,11.200,0.0000,0.0000,-170.0000
C00616=20.250,30.500,11.200,0.0000,0.0000,-170.0000
C00617=20.250,25.500,11.200,0.0000,0.0000,-170.0000
C00618=20.250,20.500,11.200,0.0000,0.0000,-170.0000
C00619=20.250,15.500,11.200,0.0000,0.0000,-170.0000
C00620=20.250,10.500,11.200,0.0000,0.0000,-170.0000
C00621=20.250,5.500,11.200,0.0000,0.0000,-170.0000
C00622=20.250,0.500,11.200,0.0000,0.0000,-170.0000
C00623=20.250,-4.500,11.200,0.0000,0.0000,-170.0000
C00624=20.250,-9.500,11.200,0.0000,0.0000,-170.0000
C00625=20.250,-14.500,11.200,0.0000,0.0000,-170.0000
C00626=20.250,-19.500,11.200,0.0000,0.0000,-170.0000
C00627=20.250,-24.500,11.200,0.0000,0.0000,-170.0000
C00628=20.250,-29.500,11.200,0.0000,0.0000,-170.0000
C00629=15.525,-29.500,11.200,0.0000,0.0000,-170.0000
C00630=10.800,-29.500,11.200,0.0000,0.0000,-170.0000
C00631=6.075,-29.500,11.200,0.0000,0.0000,-170.0000
C00632=1.350,-29.500,11.200,0.0000,0.0000,-170.0000
C00633=-3.375,-29.500,11.200,0.0000,0.0000,-170.0000
C00634=-8.100,-29.500,11.200,0.0000,0.0000,-170.0000
C00635=-12.825,-29.500,11.200,0.0000,0.0000,-170.0000
C00636=-17.550,-29.500,11.200,0.0000,0.0000,-170.0000
C00637=-22.275,-29.500,11.200,0.0000,0.0000,-170.0000
C00638=-27.000,-29.500,11.200,0.0000,0.0000,-170.0000
C00639=-27.000,-29.500,12.900,0.0000,0.0000,-170.0000
C00640=-22.275,-29.500,12.900,0.0000,0.0000,-170.0000
C00641=-17.550,-29.500,12.900,0.0000,0.0000,-170.0000
C00642=-12.825,-29.500,12.900,0.0000,0.0000,-170.0000
C00643=-8.100,-29.500,12.900,0.0000,0.0000,-170.0000
C00644=-3.375,-29.500,12.900,0.0000,0.0000,-170.0000
C00645=1.350,-29.500,12.900,0.0000,0.0000,-170.0000
C00646=6.075,-29.500,12.900,0.0000,0.0000,-170.0000
C00647=10.800,-29.500,12.900,0.0000,0.0000,-170.0000
C00648=15.525,-29.500,12.900,0.0000,0.0000,-170.0000
C00649=20.250,-29.500,12.900,0.0000,0.0000,-170.0000
C00650=20.250,-24.500,12.900,0.0000,0.0000,-170.0000
C00651=20.250,-19.500,12.900,0.0000,0.0000,-170.0000
C00652=20.250,-14.500,12.900,0.0000,0.0000,-170.0000
C00653=20.250,-9.500,12.900,0.0000,0.0000,-170.0000
C00654=20.250,-4.500,12.900,0.0000,0.0000,-170.0000
C00655=20.250,0.500,12.900,0.0000,0.0000,-170.0000
C00656=20.250,5.500,12.900,0.0000,0.0000,-170.0000
C00657=20.250,10.500,12.900,0.0000,0.0000,-170.0000
C00658=20.250,15.500,12.900,0.0000,0.0000,-170.0000
C00659=20.250,20.500,12.900,0.0000,0.0000,-170.0000
C00660=20.250,25.500,12.900,0.0000,0.0000,-170.0000
C00661=20.250,30.500,12.900,0.0000,0.0000,-170.0000
C00662=20.250,35.500,12.900,0.0000,0.0000,-170.0000
C00663=20.250,40.500,12.900,0.0000,0.0000,-170.0000
C00664=20.250,45.500,12.900,0.0000,0.0000,-170.0000
C00665=20.250,50.500,12.900,0.0000,0.0000,-170.0000
C00666=20.250,55.500,12.900,0.0000,0.0000,-170.0000
C00667=20.250,60.500,12.900,0.0000,0.0000,-170.0000
C00668=20.250,65.500,12.900,0.0000,0.0000,-170.0000
C00669=20.250,70.500,12.900,0.0000,0.0000,-170.0000
C00670=20.250,75.500,12.900,0.0000,0.0000,-170.0000
C00671=20.250,80.500,12.900,0.0000,0.0000,-170.0000
C00672=20.250,80.500,12.900,0.0000,0.0000,-170.0000
C00673=23.000,83.250,12.900,0.0000,0.0000,-170.0000
C00674=25.750,80.500,12.900,0.0000,0.0000,-170.0000
C00675=25.750,75.500,12.900,0.0000,0.0000,-170.0000
C00676=25.750,70.500,12.900,0.0000,0.0000,-170.0000
C00677=25.750,65.500,12.900,0.0000,0.0000,-170.0000
C00678=25.750,60.500,12.900,0.0000,0.0000,-170.0000
C00679=25.750,55.500,12.900,0.0000,0.0000,-170.0000
C00680=25.750,50.500,12.900,0.0000,0.0000,-170.0000
C00681=25.750,45.500,12.900,0.0000,0.0000,-170.0000
C00682=25.750,40.500,12.900,0.0000,0.0000,-170.0000
C00683=25.750,35.500,12.900,0.0000,0.0000,-170.0000
C00684=25.750,30.500,12.900,0.0000,0.0000,-170.0000
C00685=25.750,25.500,12.900,0.0000,0.0000,-170.0000
C00686=25.750,20.500,12.900,0.0000,0.0000,-170.0000
C00687=25.750,15.500,12.900,0.0000,0.0000,-170.0000
C00688=25.750,10.500,12.900,0.0000,0.0000,-170.0000
C00689=25.750,5.500,12.900,0.0000,0.0000,-170.0000
C00690=25.750,0.500,12.900,0.0000,0.0000,-170.0000
C00691=25.750,-4.500,12.900,0.0000,0.0000,-170.0000
C00692=25.750,-9.500,12.900,0.0000,0.0000,-170.0000
C00693=25.750,-14.500,12.900,0.0000,0.0000,-170.0000
C00694=25.750,-19.500,12.900,0.0000,0.0000,-170.0000
C00695=25.750,-24.500,12.900,0.0000,0.0000,-170.0000
C00696=25.750,-29.500,12.900,0.0000,0.0000,-170.0000
C00697=30.475,-29.500,12.900,0.0000,0.0000,-170.0000
C00698=35.200,-29.500,12.900,0.0000,0.0000,-170.0000
C00699=39.925,-29.500,12.900,0.0000,0.0000,-170.0000
C00700=44.650,-29.500,12.900,0.0000,0.0000,-170.0000
C00701=49.375,-29.500,12.900,0.0000,0.0000,-170.0000
C00702=54.100,-29.500,12.900,0.0000,0.0000,-170.0000
C00703=58.825,-29.500,12.900,0.0000,0.0000,-170.0000
C00704=63.550,-29.500,12.900,0.0000,0.0000,-170.0000
C00705=68.275,-29.500,12.900,0.0000,0.0000,-170.0000
C00706=73.000,-29.500,12.900,0.0000,0.0000,-170.0000
C00707=73.000,-29.500,12.900,0.0000,0.0000,-170.0000
C00708=75.750,-32.250,12.900,0.0000,0.0000,-170.0000
C00709=73.000,-35.000,12.900,0.0000,0.0000,-170.0000
C00710=68.000,-35.000,12.900,0.0000,0.0000,-170.0000
C00711=63.000,-35.000,12.900,0.0000,0.0000,-170.0000
C00712=58.000,-35.000,12.900,0.0000,0.0000,-170.0000
C00713=53.000,-35.000,12.900,0.0000,0.0000,-170.0000
C00714=48.000,-35.000,12.900,0.0000,0.0000,-170.0000
C00715=43.000,-35.000,12.900,0.0000,0.0000,-170.0000
C00716=38.000,-35.000,12.900,0.0000,0.0000,-170.0000
C00717=33.000,-35.000,12.900,0.0000,0.0000,-170.0000
C00718=28.000,-35.000,12.900,0.0000,0.0000,-170.0000
C00719=23.000,-35.000,12.900,0.0000,0.0000,-170.0000
C00720=18.000,-35.000,12.900,0.0000,0.0000,-170.0000
C00721=13.000,-35.000,12.900,0.0000,0.0000,-170.0000
C00722=8.000,-35.000,12.900,0.0000,0.0000,-170.0000
C00723=3.000,-35.000,12.900,0.0000,0.0000,-170.0000
C00724=-2.000,-35.000,12.900,0.0000,0.0000,-170.0000
C00725=-7.000,-35.000,12.900,0.0000,0.0000,-170.0000
C00726=-12.000,-35.000,12.900,0.0000,0.0000,-170.0000
C00727=-17.000,-35.000,12.900,0.0000,0.0000,-170.0000
C00728=-22.000,-35.000,12.900,0.0000,0.0000,-170.0000
C00729=-27.000,-35.000,12.900,0.0000,0.0000,-170.0000
C00730=-27.000,-35.000,14.600,0.0000,0.0000,-170.0000
C00731=-22.000,-35.000,14.600,0.0000,0.0000,-170.0000
C00732=-17.000,-35.000,14.600,0.0000,0.0000,-170.0000
C00733=-12.000,-35.000,14.600,0.0000,0.0000,-170.0000
C00734=-7.000,-35.000,14.600,0.0000,0.0000,-170.0000
C00735=-2.000,-35.000,14.600,0.0000,0.0000,-170.0000
C00736=3.000,-35.000,14.600,0.0000,0.0000,-170.0000
C00737=8.000,-35.000,14.600,0.0000,0.0000,-170.0000
C00738=13.000,-35.000,14.600,0.0000,0.0000,-170.0000
C00739=18.000,-35.000,14.600,0.0000,0.0000,-170.0000
C00740=23.000,-35.000,14.600,0.0000,0.0000,-170.0000
C00741=28.000,-35.000,14.600,0.0000,0.0000,-170.0000
C00742=33.000,-35.000,14.600,0.0000,0.0000,-170.0000
C00743=38.000,-35.000,14.600,0.0000,0.0000,-170.0000
C00744=43.000,-35.000,14.600,0.0000,0.0000,-170.0000
C00745=48.000,-35.000,14.600,0.0000,0.0000,-170.0000
C00746=53.000,-35.000,14.600,0.0000,0.0000,-170.0000
C00747=58.000,-35.000,14.600,0.0000,0.0000,-170.0000
C00748=63.000,-35.000,14.600,0.0000,0.0000,-170.0000
C00749=68.000,-35.000,14.600,0.0000,0.0000,-170.0000
C00750=73.000,-35.000,14.600,0.0000,0.0000,-170.0000
C00751=73.000,-35.000,14.600,0.0000,0.0000,-170.0000
C00752=75.750,-32.250,14.600,0.0000,0.0000,-170.0000
C00753=73.000,-29.500,14.600,0.0000,0.0000,-170.0000
C00754=68.275,-29.500,14.600,0.0000,0.0000,-170.0000
C00755=63.550,-29.500,14.600,0.0000,0.0000,-170.0000
C00756=58.825,-29.500,14.600,0.0000,0.0000,-170.0000
C00757=54.100,-29.500,14.600,0.0000,0.0000,-170.0000
C00758=49.375,-29.500,14.600,0.0000,0.0000,-170.0000
C00759=44.650,-29.500,14.600,0.0000,0.0000,-170.0000
C00760=39.925,-29.500,14.600,0.0000,0.0000,-170.0000
C00761=35.200,-29.500,14.600,0.0000,0.0000,-170.0000
C00762=30.475,-29.500,14.600,0.0000,0.0000,-170.0000
C00763=25.750,-29.500,14.600,0.0000,0.0000,-170.0000
C00764=25.750,-24.500,14.600,0.0000,0.0000,-170.0000
C00765=25.750,-19.500,14.600,0.0000,0.0000,-170.0000
C00766=25.750,-14.500,14.600,0.0000,0.0000,-170.0000
C00767=25.750,-9.500,14.600,0.0000,0.0000,-170.0000
C00768=25.750,-4.500,14.600,0.0000,0.0000,-170.0000
C00769=25.750,0.500,14.600,0.0000,0.0000,-170.0000
C00770=25.750,5.500,14.600,0.0000,0.0000,-170.0000
C00771=25.750,10.500,14.600,0.0000,0.0000,-170.0000
C00772=25.750,15.500,14.600,0.0000,0.0000,-170.0000
C00773=25.750,20.500,14.600,0.0000,0.0000,-170.0000
C00774=25.750,25.500,14.600,0.0000,0.0000,-170.0000
C00775=25.750,30.500,14.600,0.0000,0.0000,-170.0000
C00776=25.750,35.500,14.600,0.0000,0.0000,-170.0000
C00777=25.750,40.500,14.600,0.0000,0.0000,-170.0000
C00778=25.750,45.500,14.600,0.0000,0.0000,-170.0000
C00779=25.750,50.500,14.600,0.0000,0.0000,-170.0000
C00780=25.750,55.500,14.600,0.0000,0.0000,-170.0000
C00781=25.750,60.500,14.600,0.0000,0.0000,-170.0000
C00782=25.750,65.500,14.600,0.0000,0.0000,-170.0000
C00783=25.750,70.500,14.600,0.0000,0.0000,-170.0000
C00784=25.750,75.500,14.600,0.0000,0.0000,-170.0000
C00785=25.750,80.500,14.600,0.0000,0.0000,-170.0000
C00786=25.750,80.500,14.600,0.0000,0.0000,-170.0000
C00787=23.000,83.250,14.600,0.0000,0.0000,-170.0000
C00788=20.250,80.500,14.600,0.0000,0.0000,-170.0000
C00789=20.250,75.500,14.600,0.0000,0.0000,-170.0000
C00790=20.250,70.500,14.600,0.0000,0.0000,-170.0000
C00791=20.250,65.500,14.600,0.0000,0.0000,-170.0000
C00792=20.250,60.500,14.600,0.0000,0.0000,-170.0000
C00793=20.250,55.500,14.600,0.0000,0.0000,-170.0000
C00794=20.250,50.500,14.600,0.0000,0.0000,-170.0000
C00795=20.250,45.500,14.600,0.0000,0.0000,-170.0000
C00796=20.250,40.500,14.600,0.0000,0.0000,-170.0000
C00797=20.250,35.500,14.600,0.0000,0.0000,-170.0000
C00798=20.250,30.500,14.600,0.0000,0.0000,-170.0000
C00799=20.250,25.500,14.600,0.0000,0.0000,-170.0000
C00800=20.250,20.500,14.600,0.0000,0.0000,-170.0000
C00801=20.250,15.500,14.600,0.0000,0.0000,-170.0000
C00802=20.250,10.500,14.600,0.0000,0.0000,-170.0000
C00803=20.250,5.500,14.600,0.0000,0.0000,-170.0000
C00804=20.250,0.500,14.600,0.0000,0.0000,-170.0000
C00805=20.250,-4.500,14.600,0.0000,0.0000,-170.0000
C00806=20.250,-9.500,14.600,0.0000,0.0000,-170.0000
C00807=20.250,-14.500,14.600,0.0000,0.0000,-170.0000
C00808=20.250,-19.500,14.600,0.0000,0.0000,-170.0000
C00809=20.250,-24.500,14.600,0.0000,0.0000,-170.0000
C00810=20.250,-29.500,14.600,0.0000,0.0000,-170.0000
C00811=15.525,-29.500,14.600,0.0000,0.0000,-170.0000
C00812=10.800,-29.500,14.600,0.0000,0.0000,-170.0000
C00813=6.075,-29.500,14.600,0.0000,0.0000,-170.0000
C00814=1.350,-29.500,14.600,0.0000,0.0000,-170.0000
C00815=-3.375,-29.500,14.600,0.0000,0.0000,-170.0000
C00816=-8.100,-29.500,14.600,0.0000,0.0000,-170.0000
C00817=-12.825,-29.500,14.600,0.0000,0.0000,-170.0000
C00818=-17.550,-29.500,14.600,0.0000,0.0000,-170.0000
C00819=-22.275,-29.500,14.600,0.0000,0.0000,-170.0000
C00820=-27.000,-29.500,14.600,0.0000,0.0000,-170.0000
C00821=-27.000,-29.500,16.300,0.0000,0.0000,-170.0000
C00822=-22.275,-29.500,16.300,0.0000,0.0000,-170.0000
C00823=-17.550,-29.500,16.300,0.0000,0.0000,-170.0000
C00824=-12.825,-29.500,16.300,0.0000,0.0000,-170.0000
C00825=-8.100,-29.500,16.300,0.0000,0.0000,-170.0000
C00826=-3.375,-29.500,16.300,0.0000,0.0000,-170.0000
C00827=1.350,-29.500,16.300,0.0000,0.0000,-170.0000
C00828=6.075,-29.500,16.300,0.0000,0.0000,-170.0000
C00829=10.800,-29.500,16.300,0.0000,0.0000,-170.0000
C00830=15.525,-29.500,16.300,0.0000,0.0000,-170.0000
C00831=20.250,-29.500,16.300,0.0000,0.0000,-170.0000
C00832=20.250,-24.500,16.300,0.0000,0.0000,-170.0000
C00833=20.250,-19.500,16.300,0.0000,0.0000,-170.0000
C00834=20.250,-14.500,16.300,0.0000,0.0000,-170.0000
C00835=20.250,-9.500,16.300,0.0000,0.0000,-170.0000
C00836=20.250,-4.500,16.300,0.0000,0.0000,-170.0000
C00837=20.250,0.500,16.300,0.0000,0.0000,-170.0000
C00838=20.250,5.500,16.300,0.0000,0.0000,-170.0000
C00839=20.250,10.500,16.300,0.0000,0.0000,-170.0000
C00840=20.250,15.500,16.300,0.0000,0.0000,-170.0000
C00841=20.250,20.500,16.300,0.0000,0.0000,-170.0000
C00842=20.250,25.500,16.300,0.0000,0.0000,-170.0000
C00843=20.250,30.500,16.300,0.0000,0.0000,-170.0000
C00844=20.250,35.500,16.300,0.0000,0.0000,-170.0000
C00845=20.250,40.500,16.300,0.0000,0.0000,-170.0000
C00846=20.250,45.500,16.300,0.0000,0.0000,-170.0000
C00847=20.250,50.500,16.300,0.0000,0.0000,-170.0000
C00848=20.250,55.500,16.300,0.0000,0.0000,-170.0000
C00849=20.250,60.500,16.300,0.0000,0.0000,-170.0000
C00850=20.250,65.500,16.300,0.0000,0.0000,-170.0000
C00851=20.250,70.500,16.300,0.0000,0.0000,-170.0000
C00852=20.250,75.500,16.300,0.0000,0.0000,-170.0000
C00853=20.250,80.500,16.300,0.0000,0.0000,-170.0000
C00854=20.250,80.500,16.300,0.0000,0.0000,-170.0000
C00855=23.000,83.250,16.300,0.0000,0.0000,-170.0000
C00856=25.750,80.500,16.300,0.0000,0.0000,-170.0000
C00857=25.750,75.500,16.300,0.0000,0.0000,-170.0000
C00858=25.750,70.500,16.300,0.0000,0.0000,-170.0000
C00859=25.750,65.500,16.300,0.0000,0.0000,-170.0000
C00860=25.750,60.500,16.300,0.0000,0.0000,-170.0000
C00861=25.750,55.500,16.300,0.0000,0.0000,-170.0000
C00862=25.750,50.500,16.300,0.0000,0.0000,-170.0000
C00863=25.750,45.500,16.300,0.0000,0.0000,-170.0000
C00864=25.750,40.500,16.300,0.0000,0.0000,-170.0000
C00865=25.750,35.500,16.300,0.0000,0.0000,-170.0000
C00866=25.750,30.500,16.300,0.0000,0.0000,-170.0000
C00867=25.750,25.500,16.300,0.0000,0.0000,-170.0000
C00868=25.750,20.500,16.300,0.0000,0.0000,-170.0000
C00869=25.750,15.500,16.300,0.0000,0.0000,-170.0000
C00870=25.750,10.500,16.300,0.0000,0.0000,-170.0000
C00871=25.750,5.500,16.300,0.0000,0.0000,-170.0000
C00872=25.750,0.500,16.300,0.0000,0.0000,-170.0000
C00873=25.750,-4.500,16.300,0.0000,0.0000,-170.0000
C00874=25.750,-9.500,16.300,0.0000,0.0000,-170.0000
C00875=25.750,-14.500,16.300,0.0000,0.0000,-170.0000
C00876=25.750,-19.500,16.300,0.0000,0.0000,-170.0000
C00877=25.750,-24.500,16.300,0.0000,0.0000,-170.0000
C00878=25.750,-29.500,16.300,0.0000,0.0000,-170.0000
C00879=30.475,-29.500,16.300,0.0000,0.0000,-170.0000
C00880=35.200,-29.500,16.300,0.0000,0.0000,-170.0000
C00881=39.925,-29.500,16.300,0.0000,0.0000,-170.0000
C00882=44.650,-29.500,16.300,0.0000,0.0000,-170.0000
C00883=49.375,-29.500,16.300,0.0000,0.0000,-170.0000
C00884=54.100,-29.500,16.300,0.0000,0.0000,-170.0000
C00885=58.825,-29.500,16.300,0.0000,0.0000,-170.0000
C00886=63.550,-29.500,16.300,0.0000,0.0000,-170.0000
C00887=68.275,-29.500,16.300,0.0000,0.0000,-170.0000
C00888=73.000,-29.500,16.300,0.0000,0.0000,-170.0000
C00889=73.000,-29.500,16.300,0.0000,0.0000,-170.0000
C00890=75.750,-32.250,16.300,0.0000,0.0000,-170.0000
C00891=73.000,-35.000,16.300,0.0000,0.0000,-170.0000
C00892=68.000,-35.000,16.300,0.0000,0.0000,-170.0000
C00893=63.000,-35.000,16.300,0.0000,0.0000,-170.0000
C00894=58.000,-35.000,16.300,0.0000,0.0000,-170.0000
C00895=53.000,-35.000,16.300,0.0000,0.0000,-170.0000
C00896=48.000,-35.000,16.300,0.0000,0.0000,-170.0000
C00897=43.000,-35.000,16.300,0.0000,0.0000,-170.0000
C00898=38.000,-35.000,16.300,0.0000,0.0000,-170.0000
C00899=33.000,-35.000,16.300,0.0000,0.0000,-170.0000
C00900=28.000,-35.000,16.300,0.0000,0.0000,-170.0000
C00901=23.000,-35.000,16.300,0.0000,0.0000,-170.0000
C00902=18.000,-35.000,16.300,0.0000,0.0000,-170.0000
C00903=13.000,-35.000,16.300,0.0000,0.0000,-170.0000
C00904=8.000,-35.000,16.300,0.0000,0.0000,-170.0000
C00905=3.000,-35.000,16.300,0.0000,0.0000,-170.0000
C00906=-2.000,-35.000,16.300,0.0000,0.0000,-170.0000
C00907=-7.000,-35.000,16.300,0.0000,0.0000,-170.0000
C00908=-12.000,-35.000,16.300,0.0000,0.0000,-170.0000
C00909=-17.000,-35.000,16.300,0.0000,0.0000,-170.0000
C00910=-22.000,-35.000,16.300,0.0000,0.0000,-170.0000
C00911=-27.000,-35.000,16.300,0.0000,0.0000,-170.0000
C00912=-27.000,-35.000,18.000,0.0000,0.0000,-170.0000
C00913=-22.000,-35.000,18.000,0.0000,0.0000,-170.0000
C00914=-17.000,-35.000,18.000,0.0000,0.0000,-170.0000
C00915=-12.000,-35.000,18.000,0.0000,0.0000,-170.0000
C00916=-7.000,-35.000,18.000,0.0000,0.0000,-170.0000
C00917=-2.000,-35.000,18.000,0.0000,0.0000,-170.0000
C00918=3.000,-35.000,18.000,0.0000,0.0000,-170.0000
C00919=8.000,-35.000,18.000,0.0000,0.0000,-170.0000
C00920=13.000,-35.000,18.000,0.0000,0.0000,-170.0000
C00921=18.000,-35.000,18.000,0.0000,0.0000,-170.0000
C00922=23.000,-35.000,18.000,0.0000,0.0000,-170.0000
C00923=28.000,-35.000,18.000,0.0000,0.0000,-170.0000
C00924=33.000,-35.000,18.000,0.0000,0.0000,-170.0000
C00925=38.000,-35.000,18.000,0.0000,0.0000,-170.0000
C00926=43.000,-35.000,18.000,0.0000,0.0000,-170.0000
C00927=48.000,-35.000,18.000,0.0000,0.0000,-170.0000
C00928=53.000,-35.000,18.000,0.0000,0.0000,-170.0000
C00929=58.000,-35.000,18.000,0.0000,0.0000,-170.0000
C00930=63.000,-35.000,18.000,0.0000,0.0000,-170.0000
C00931=68.000,-35.000,18.000,0.0000,0.0000,-170.0000
C00932=73.000,-35.000,18.000,0.0000,0.0000,-170.0000
C00933=73.000,-35.000,18.000,0.0000,0.0000,-170.0000
C00934=75.750,-32.250,18.000,0.0000,0.0000,-170.0000
C00935=73.000,-29.500,18.000,0.0000,0.0000,-170.0000
C00936=68.275,-29.500,18.000,0.0000,0.0000,-170.0000
C00937=63.550,-29.500,18.000,0.0000,0.0000,-170.0000
C00938=58.825,-29.500,18.000,0.0000,0.0000,-170.0000
C00939=54.100,-29.500,18.000,0.0000,0.0000,-170.0000
C00940=49.375,-29.500,18.000,0.0000,0.0000,-170.0000
C00941=44.650,-29.500,18.000,0.0000,0.0000,-170.0000
C00942=39.925,-29.500,18.000,0.0000,0.0000,-170.0000
C00943=35.200,-29.500,18.000,0.0000,0.0000,-170.0000
C00944=30.475,-29.500,18.000,0.0000,0.0000,-170.0000
C00945=25.750,-29.500,18.000,0.0000,0.0000,-170.0000
C00946=25.750,-24.500,18.000,0.0000,0.0000,-170.0000
C00947=25.750,-19.500,18.000,0.0000,0.0000,-170.0000
C00948=25.750,-14.500,18.000,0.0000,0.0000,-170.0000
C00949=25.750,-9.500,18.000,0.0000,0.0000,-170.0000
C00950=25.750,-4.500,18.000,0.0000,0.0000,-170.0000
C00951=25.750,0.500,18.000,0.0000,0.0000,-170.0000
C00952=25.750,5.500,18.000,0.0000,0.0000,-170.0000
C00953=25.750,10.500,18.000,0.0000,0.0000,-170.0000
C00954=25.750,15.500,18.000,0.0000,0.0000,-170.0000
C00955=25.750,20.500,18.000,0.0000,0.0000,-170.0000
C00956=25.750,25.500,18.000,0.0000,0.0000,-170.0000
C00957=25.750,30.500,18.000,0.0000,0.0000,-170.0000
C00958=25.750,35.500,18.000,0.0000,0.0000,-170.0000
C00959=25.750,40.500,18.000,0.0000,0.0000,-170.0000
C00960=25.750,45.500,18.000,0.0000,0.0000,-170.0000
C00961=25.750,50.500,18.000,0.0000,0.0000,-170.0000
C00962=25.750,55.500,18.000,0.0000,0.0000,-170.0000
C00963=25.750,60.500,18.000,0.0000,0.0000,-170.0000
C00964=25.750,65.500,18.000,0.0000,0.0000,-170.0000
C00965=25.750,70.500,18.000,0.0000,0.0000,-170.0000
C00966=25.750,75.500,18.000,0.0000,0.0000,-170.0000
C00967=25.750,80.500,18.000,0.0000,0.0000,-170.0000
C00968=25.750,80.500,18.000,0.0000,0.0000,-170.0000
C00969=23.000,83.250,18.000,0.0000,0.0000,-170.0000
C00970=20.250,80.500,18.000,0.0000,0.0000,-170.0000
C00971=20.250,75.500,18.000,0.0000,0.0000,-170.0000
C00972=20.250,70.500,18.000,0.0000,0.0000,-170.0000
C00973=20.250,65.500,18.000,0.0000,0.0000,-170.0000
C00974=20.250,60.500,18.000,0.0000,0.0000,-170.0000
C00975=20.250,55.500,18.000,0.0000,0.0000,-170.0000
C00976=20.250,50.500,18.000,0.0000,0.0000,-170.0000
C00977=20.250,45.500,18.000,0.0000,0.0000,-170.0000
C00978=20.250,40.500,18.000,0.0000,0.0000,-170.0000
C00979=20.250,35.500,18.000,0.0000,0.0000,-170.0000
C00980=20.250,30.500,18.000,0.0000,0.0000,-170.0000
C00981=20.250,25.500,18.000,0.0000,0.0000,-170.0000
C00982=20.250,20.500,18.000,0.0000,0.0000,-170.0000
C00983=20.250,15.500,18.000,0.0000,0.0000,-170.0000
C00984=20.250,10.500,18.000,0.0000,0.0000,-170.0000
C00985=20.250,5.500,18.000,0.0000,0.0000,-170.0000
C00986=20.250,0.500,18.000,0.0000,0.0000,-170.0000
C00987=20.250,-4.500,18.000,0.0000,0.0000,-170.0000
C00988=20.250,-9.500,18.000,0.0000,0.0000,-170.0000
C00989=20.250,-14.500,18.000,0.0000,0.0000,-170.0000
C00990=20.250,-19.500,18.000,0.0000,0.0000,-170.0000
C00991=20.250,-24.500,18.000,0.0000,0.0000,-170.0000
C00992=20.250,-29.500,18.000,0.0000,0.0000,-170.0000
C00993=15.525,-29.500,18.000,0.0000,0.0000,-170.0000
C00994=10.800,-29.500,18.000,0.0000,0.0000,-170.0000
C00995=6.075,-29.500,18.000,0.0000,0.0000,-170.0000
C00996=1.350,-29.500,18.000,0.0000,0.0000,-170.0000
C00997=-3.375,-29.500,18.000,0.0000,0.0000,-170.0000
C00998=-8.100,-29.500,18.000,0.0000,0.0000,-170.0000
C00999=-12.825,-29.500,18.000,0.0000,0.0000,-170.0000
C01000=-17.550,-29.500,18.000,0.0000,0.0000,-170.0000
C01001=-22.275,-29.500,18.000,0.0000,0.0000,-170.0000
C01002=-27.000,-29.500,18.000,0.0000,0.0000,-170.0000
C01003=-27.000,-29.500,19.700,0.0000,0.0000,-170.0000
C01004=-22.275,-29.500,19.700,0.0000,0.0000,-170.0000
C01005=-17.550,-29.500,19.700,0.0000,0.0000,-170.0000
C01006=-12.825,-29.500,19.700,0.0000,0.0000,-170.0000
C01007=-8.100,-29.500,19.700,0.0000,0.0000,-170.0000
C01008=-3.375,-29.500,19.700,0.0000,0.0000,-170.0000
C01009=1.350,-29.500,19.700,0.0000,0.0000,-170.0000
C01010=6.075,-29.500,19.700,0.0000,0.0000,-170.0000
C01011=10.800,-29.500,19.700,0.0000,0.0000,-170.0000
C01012=15.525,-29.500,19.700,0.0000,0.0000,-170.0000
C01013=20.250,-29.500,19.700,0.0000,0.0000,-170.0000
C01014=20.250,-24.500,19.700,0.0000,0.0000,-170.0000
C01015=20.250,-19.500,19.700,0.0000,0.0000,-170.0000
C01016=20.250,-14.500,19.700,0.0000,0.0000,-170.0000
C01017=20.250,-9.500,19.700,0.0000,0.0000,-170.0000
C01018=20.250,-4.500,19.700,0.0000,0.0000,-170.0000
C01019=20.250,0.500,19.700,0.0000,0.0000,-170.0000
C01020=20.250,5.500,19.700,0.0000,0.0000,-170.0000
C01021=20.250,10.500,19.700,0.0000,0.0000,-170.0000
C01022=20.250,15.500,19.700,0.0000,0.0000,-170.0000
C01023=20.250,20.500,19.700,0.0000,0.0000,-170.0000
C01024=20.250,25.500,19.700,0.0000,0.0000,-170.0000
C01025=20.250,30.500,19.700,0.0000,0.0000,-170.0000
C01026=20.250,35.500,19.700,0.0000,0.0000,-170.0000
C01027=20.250,40.500,19.700,0.0000,0.0000,-170.0000
C01028=20.250,45.500,19.700,0.0000,0.0000,-170.0000
C01029=20.250,50.500,19.700,0.0000,0.0000,-170.0000
C01030=20.250,55.500,19.700,0.0000,0.0000,-170.0000
C01031=20.250,60.500,19.700,0.0000,0.0000,-170.0000
C01032=20.250,65.500,19.700,0.0000,0.0000,-170.0000
C01033=20.250,70.500,19.700,0.0000,0.0000,-170.0000
C01034=20.250,75.500,19.700,0.0000,0.0000,-170.0000
C01035=20.250,80.500,19.700,0.0000,0.0000,-170.0000
C01036=20.250,80.500,19.700,0.0000,0.0000,-170.0000
C01037=23.000,83.250,19.700,0.0000,0.0000,-170.0000
C01038=25.750,80.500,19.700,0.0000,0.0000,-170.0000
C01039=25.750,75.500,19.700,0.0000,0.0000,-170.0000
C01040=25.750,70.500,19.700,0.0000,0.0000,-170.0000
C01041=25.750,65.500,19.700,0.0000,0.0000,-170.0000
C01042=25.750,60.500,19.700,0.0000,0.0000,-170.0000
C01043=25.750,55.500,19.700,0.0000,0.0000,-170.0000
C01044=25.750,50.500,19.700,0.0000,0.0000,-170.0000
C01045=25.750,45.500,19.700,0.0000,0.0000,-170.0000
C01046=25.750,40.500,19.700,0.0000,0.0000,-170.0000
C01047=25.750,35.500,19.700,0.0000,0.0000,-170.0000
C01048=25.750,30.500,19.700,0.0000,0.0000,-170.0000
C01049=25.750,25.500,19.700,0.0000,0.0000,-170.0000
C01050=25.750,20.500,19.700,0.0000,0.0000,-170.0000
C01051=25.750,15.500,19.700,0.0000,0.0000,-170.0000
C01052=25.750,10.500,19.700,0.0000,0.0000,-170.0000
C01053=25.750,5.500,19.700,0.0000,0.0000,-170.0000
C01054=25.750,0.500,19.700,0.0000,0.0000,-170.0000
C01055=25.750,-4.500,19.700,0.0000,0.0000,-170.0000
C01056=25.750,-9.500,19.700,0.0000,0.0000,-170.0000
C01057=25.750,-14.500,19.700,0.0000,0.0000,-170.0000
C01058=25.750,-19.500,19.700,0.0000,0.0000,-170.0000
C01059=25.750,-24.500,19.700,0.0000,0.0000,-170.0000
C01060=25.750,-29.500,19.700,0.0000,0.0000,-170.0000
C01061=30.475,-29.500,19.700,0.0000,0.0000,-170.0000
C01062=35.200,-29.500,19.700,0.0000,0.0000,-170.0000
C01063=39.925,-29.500,19.700,0.0000,0.0000,-170.0000
C01064=44.650,-29.500,19.700,0.0000,0.0000,-170.0000
C01065=49.375,-29.500,19.700,0.0000,0.0000,-170.0000
C01066=54.100,-29.500,19.700,0.0000,0.0000,-170.0000
C01067=58.825,-29.500,19.700,0.0000,0.0000,-170.0000
C01068=63.550,-29.500,19.700,0.0000,0.0000,-170.0000
C01069=68.275,-29.500,19.700,0.0000,0.0000,-170.0000
C01070=73.000,-29.500,19.700,0.0000,0.0000,-170.0000
C01071=73.000,-29.500,19.700,0.0000,0.0000,-170.0000
C01072=75.750,-32.250,19.700,0.0000,0.0000,-170.0000
C01073=73.000,-35.000,19.700,0.0000,0.0000,-170.0000
C01074=68.000,-35.000,19.700,0.0000,0.0000,-170.0000
C01075=63.000,-35.000,19.700,0.0000,0.0000,-170.0000
C01076=58.000,-35.000,19.700,0.0000,0.0000,-170.0000
C01077=53.000,-35.000,19.700,0.0000,0.0000,-170.0000
C01078=48.000,-35.000,19.700,0.0000,0.0000,-170.0000
C01079=43.000,-35.000,19.700,0.0000,0.0000,-170.0000
C01080=38.000,-35.000,19.700,0.0000,0.0000,-170.0000
C01081=33.000,-35.000,19.700,0.0000,0.0000,-170.0000
C01082=28.000,-35.000,19.700,0.0000,0.0000,-170.0000
C01083=23.000,-35.000,19.700,0.0000,0.0000,-170.0000
C01084=18.000,-35.000,19.700,0.0000,0.0000,-170.0000
C01085=13.000,-35.000,19.700,0.0000,0.0000,-170.0000
C01086=8.000,-35.000,19.700,0.0000,0.0000,-170.0000
C01087=3.000,-35.000,19.700,0.0000,0.0000,-170.0000
C01088=-2.000,-35.000,19.700,0.0000,0.0000,-170.0000
C01089=-7.000,-35.000,19.700,0.0000,0.0000,-170.0000
C01090=-12.000,-35.000,19.700,0.0000,0.0000,-170.0000
C01091=-17.000,-35.000,19.700,0.0000,0.0000,-170.0000
C01092=-22.000,-35.000,19.700,0.0000,0.0000,-170.0000
C01093=-27.000,-35.000,19.700,0.0000,0.0000,-170.0000
C01094=-27.000,-35.000,21.400,0.0000,0.0000,-170.0000
C01095=-22.000,-35.000,21.400,0.0000,0.0000,-170.0000
C01096=-17.000,-35.000,21.400,0.0000,0.0000,-170.0000
C01097=-12.000,-35.000,21.400,0.0000,0.0000,-170.0000
C01098=-7.000,-35.000,21.400,0.0000,0.0000,-170.0000
C01099=-2.000,-35.000,21.400,0.0000,0.0000,-170.0000
C01100=3.000,-35.000,21.400,0.0000,0.0000,-170.0000
C01101=8.000,-35.000,21.400,0.0000,0.0000,-170.0000
C01102=13.000,-35.000,21.400,0.0000,0.0000,-170.0000
C01103=18.000,-35.000,21.400,0.0000,0.0000,-170.0000
C01104=23.000,-35.000,21.400,0.0000,0.0000,-170.0000
C01105=28.000,-35.000,21.400,0.0000,0.0000,-170.0000
C01106=33.000,-35.000,21.400,0.0000,0.0000,-170.0000
C01107=38.000,-35.000,21.400,0.0000,0.0000,-170.0000
C01108=43.000,-35.000,21.400,0.0000,0.0000,-170.0000
C01109=48.000,-35.000,21.400,0.0000,0.0000,-170.0000
C01110=53.000,-35.000,21.400,0.0000,0.0000,-170.0000
C01111=58.000,-35.000,21.400,0.0000,0.0000,-170.0000
C01112=63.000,-35.000,21.400,0.0000,0.0000,-170.0000
C01113=68.000,-35.000,21.400,0.0000,0.0000,-170.0000
C01114=73.000,-35.000,21.400,0.0000,0.0000,-170.0000
C01115=73.000,-35.000,21.400,0.0000,0.0000,-170.0000
C01116=75.750,-32.250,21.400,0.0000,0.0000,-170.0000
C01117=73.000,-29.500,21.400,0.0000,0.0000,-170.0000
C01118=68.275,-29.500,21.400,0.0000,0.0000,-170.0000
C01119=63.550,-29.500,21.400,0.0000,0.0000,-170.0000
C01120=58.825,-29.500,21.400,0.0000,0.0000,-170.0000
C01121=54.100,-29.500,21.400,0.0000,0.0000,-170.0000
C01122=49.375,-29.500,21.400,0.0000,0.0000,-170.0000
C01123=44.650,-29.500,21.400,0.0000,0.0000,-170.0000
C01124=39.925,-29.500,21.400,0.0000,0.0000,-170.0000
C01125=35.200,-29.500,21.400,0.0000,0.0000,-170.0000
C01126=30.475,-29.500,21.400,0.0000,0.0000,-170.0000
C01127=25.750,-29.500,21.400,0.0000,0.0000,-170.0000
C01128=25.750,-24.500,21.400,0.0000,0.0000,-170.0000
C01129=25.750,-19.500,21.400,0.0000,0.0000,-170.0000
C01130=25.750,-14.500,21.400,0.0000,0.0000,-170.0000
C01131=25.750,-9.500,21.400,0.0000,0.0000,-170.0000
C01132=25.750,-4.500,21.400,0.0000,0.0000,-170.0000
C01133=25.750,0.500,21.400,0.0000,0.0000,-170.0000
C01134=25.750,5.500,21.400,0.0000,0.0000,-170.0000
C01135=25.750,10.500,21.400,0.0000,0.0000,-170.0000
C01136=25.750,15.500,21.400,0.0000,0.0000,-170.0000
C01137=25.750,20.500,21.400,0.0000,0.0000,-170.0000
C01138=25.750,25.500,21.400,0.0000,0.0000,-170.0000
C01139=25.750,30.500,21.400,0.0000,0.0000,-170.0000
C01140=25.750,35.500,21.400,0.0000,0.0000,-170.0000
C01141=25.750,40.500,21.400,0.0000,0.0000,-170.0000
C01142=25.750,45.500,21.400,0.0000,0.0000,-170.0000
C01143=25.750,50.500,21.400,0.0000,0.0000,-170.0000
C01144=25.750,55.500,21.400,0.0000,0.0000,-170.0000
C01145=25.750,60.500,21.400,0.0000,0.0000,-170.0000
C01146=25.750,65.500,21.400,0.0000,0.0000,-170.0000
C01147=25.750,70.500,21.400,0.0000,0.0000,-170.0000
C01148=25.750,75.500,21.400,0.0000,0.0000,-170.0000
C01149=25.750,80.500,21.400,0.0000,0.0000,-170.0000
C01150=25.750,80.500,21.400,0.0000,0.0000,-170.0000
C01151=23.000,83.250,21.400,0.0000,0.0000,-170.0000
C01152=20.250,80.500,21.400,0.0000,0.0000,-170.0000
C01153=20.250,75.500,21.400,0.0000,0.0000,-170.0000
C01154=20.250,70.500,21.400,0.0000,0.0000,-170.0000
C01155=20.250,65.500,21.400,0.0000,0.0000,-170.0000
C01156=20.250,60.500,21.400,0.0000,0.0000,-170.0000
C01157=20.250,55.500,21.400,0.0000,0.0000,-170.0000
C01158=20.250,50.500,21.400,0.0000,0.0000,-170.0000
C01159=20.250,45.500,21.400,0.0000,0.0000,-170.0000
C01160=20.250,40.500,21.400,0.0000,0.0000,-170.0000
C01161=20.250,35.500,21.400,0.0000,0.0000,-170.0000
C01162=20.250,30.500,21.400,0.0000,0.0000,-170.0000
C01163=20.250,25.500,21.400,0.0000,0.0000,-170.0000
C01164=20.250,20.500,21.400,0.0000,0.0000,-170.0000
C01165=20.250,15.500,21.400,0.0000,0.0000,-170.0000
C01166=20.250,10.500,21.400,0.0000,0.0000,-170.0000
C01167=20.250,5.500,21.400,0.0000,0.0000,-170.0000
C01168=20.250,0.500,21.400,0.0000,0.0000,-170.0000
C01169=20.250,-4.500,21.400,0.0000,0.0000,-170.0000
C01170=20.250,-9.500,21.400,0.0000,0.0000,-170.0000
C01171=20.250,-14.500,21.400,0.0000,0.0000,-170.0000
C01172=20.250,-19.500,21.400,0.0000,0.0000,-170.0000
C01173=20.250,-24.500,21.400,0.0000,0.0000,-170.0000
C01174=20.250,-29.500,21.400,0.0000,0.0000,-170.0000
C01175=15.525,-29.500,21.400,0.0000,0.0000,-170.0000
C01176=10.800,-29.500,21.400,0.0000,0.0000,-170.0000
C01177=6.075,-29.500,21.400,0.0000,0.0000,-170.0000
C01178=1.350,-29.500,21.400,0.0000,0.0000,-170.0000
C01179=-3.375,-29.500,21.400,0.0000,0.0000,-170.0000
C01180=-8.100,-29.500,21.400,0.0000,0.0000,-170.0000
C01181=-12.825,-29.500,21.400,0.0000,0.0000,-170.0000
C01182=-17.550,-29.500,21.400,0.0000,0.0000,-170.0000
C01183=-22.275,-29.500,21.400,0.0000,0.0000,-170.0000
C01184=-27.000,-29.500,21.400,0.0000,0.0000,-170.0000
C01185=-27.000,-29.500,23.100,0.0000,0.0000,-170.0000
C01186=-22.275,-29.500,23.100,0.0000,0.0000,-170.0000
C01187=-17.550,-29.500,23.100,0.0000,0.0000,-170.0000
C01188=-12.825,-29.500,23.100,0.0000,0.0000,-170.0000
C01189=-8.100,-29.500,23.100,0.0000,0.0000,-170.0000
C01190=-3.375,-29.500,23.100,0.0000,0.0000,-170.0000
C01191=1.350,-29.500,23.100,0.0000,0.0000,-170.0000
C01192=6.075,-29.500,23.100,0.0000,0.0000,-170.0000
C01193=10.800,-29.500,23.100,0.0000,0.0000,-170.0000
C01194=15.525,-29.500,23.100,0.0000,0.0000,-170.0000
C01195=20.250,-29.500,23.100,0.0000,0.0000,-170.0000
C01196=20.250,-24.500,23.100,0.0000,0.0000,-170.0000
C01197=20.250,-19.500,23.100,0.0000,0.0000,-170.0000
C01198=20.250,-14.500,23.100,0.0000,0.0000,-170.0000
C01199=20.250,-9.500,23.100,0.0000,0.0000,-170.0000
C01200=20.250,-4.500,23.100,0.0000,0.0000,-170.0000
C01201=20.250,0.500,23.100,0.0000,0.0000,-170.0000
C01202=20.250,5.500,23.100,0.0000,0.0000,-170.0000
C01203=20.250,10.500,23.100,0.0000,0.0000,-170.0000
C01204=20.250,15.500,23.100,0.0000,0.0000,-170.0000
C01205=20.250,20.500,23.100,0.0000,0.0000,-170.0000
C01206=20.250,25.500,23.100,0.0000,0.0000,-170.0000
C01207=20.250,30.500,23.100,0.0000,0.0000,-170.0000
C01208=20.250,35.500,23.100,0.0000,0.0000,-170.0000
C01209=20.250,40.500,23.100,0.0000,0.0000,-170.0000
C01210=20.250,45.500,23.100,0.0000,0.0000,-170.0000
C01211=20.250,50.500,23.100,0.0000,0.0000,-170.0000
C01212=20.250,55.500,23.100,0.0000,0.0000,-170.0000
C01213=20.250,60.500,23.100,0.0000,0.0000,-170.0000
C01214=20.250,65.500,23.100,0.0000,0.0000,-170.0000
C01215=20.250,70.500,23.100,0.0000,0.0000,-170.0000
C01216=20.250,75.500,23.100,0.0000,0.0000,-170.0000
C01217=20.250,80.500,23.100,0.0000,0.0000,-170.0000
C01218=20.250,80.500,23.100,0.0000,0.0000,-170.0000
C01219=23.000,83.250,23.100,0.0000,0.0000,-170.0000
C01220=25.750,80.500,23.100,0.0000,0.0000,-170.0000
C01221=25.750,75.500,23.100,0.0000,0.0000,-170.0000
C01222=25.750,70.500,23.100,0.0000,0.0000,-170.0000
C01223=25.750,65.500,23.100,0.0000,0.0000,-170.0000
C01224=25.750,60.500,23.100,0.0000,0.0000,-170.0000
C01225=25.750,55.500,23.100,0.0000,0.0000,-170.0000
C01226=25.750,50.500,23.100,0.0000,0.0000,-170.0000
C01227=25.750,45.500,23.100,0.0000,0.0000,-170.0000
C01228=25.750,40.500,23.100,0.0000,0.0000,-170.0000
C01229=25.750,35.500,23.100,0.0000,0.0000,-170.0000
C01230=25.750,30.500,23.100,0.0000,0.0000,-170.0000
C01231=25.750,25.500,23.100,0.0000,0.0000,-170.0000
C01232=25.750,20.500,23.100,0.0000,0.0000,-170.0000
C01233=25.750,15.500,23.100,0.0000,0.0000,-170.0000
C01234=25.750,10.500,23.100,0.0000,0.0000,-170.0000
C01235=25.750,5.500,23.100,0.0000,0.0000,-170.0000
C01236=25.750,0.500,23.100,0.0000,0.0000,-170.0000
C01237=25.750,-4.500,23.100,0.0000,0.0000,-170.0000
C01238=25.750,-9.500,23.100,0.0000,0.0000,-170.0000
C01239=25.750,-14.500,23.100,0.0000,0.0000,-170.0000
C01240=25.750,-19.500,23.100,0.0000,0.0000,-170.0000
C01241=25.750,-24.500,23.100,0.0000,0.0000,-170.0000
C01242=25.750,-29.500,23.100,0.0000,0.0000,-170.0000
C01243=30.475,-29.500,23.100,0.0000,0.0000,-170.0000
C01244=35.200,-29.500,23.100,0.0000,0.0000,-170.0000
C01245=39.925,-29.500,23.100,0.0000,0.0000,-170.0000
C01246=44.650,-29.500,23.100,0.0000,0.0000,-170.0000
C01247=49.375,-29.500,23.100,0.0000,0.0000,-170.0000
C01248=54.100,-29.500,23.100,0.0000,0.0000,-170.0000
C01249=58.825,-29.500,23.100,0.0000,0.0000,-170.0000
C01250=63.550,-29.500,23.100,0.0000,0.0000,-170.0000
C01251=68.275,-29.500,23.100,0.0000,0.0000,-170.0000
C01252=73.000,-29.500,23.100,0.0000,0.0000,-170.0000
C01253=73.000,-29.500,23.100,0.0000,0.0000,-170.0000
C01254=75.750,-32.250,23.100,0.0000,0.0000,-170.0000
C01255=73.000,-35.000,23.100,0.0000,0.0000,-170.0000
C01256=68.000,-35.000,23.100,0.0000,0.0000,-170.0000
C01257=63.000,-35.000,23.100,0.0000,0.0000,-170.0000
C01258=58.000,-35.000,23.100,0.0000,0.0000,-170.0000
C01259=53.000,-35.000,23.100,0.0000,0.0000,-170.0000
C01260=48.000,-35.000,23.100,0.0000,0.0000,-170.0000
C01261=43.000,-35.000,23.100,0.0000,0.0000,-170.0000
C01262=38.000,-35.000,23.100,0.0000,0.0000,-170.0000
C01263=33.000,-35.000,23.100,0.0000,0.0000,-170.0000
C01264=28.000,-35.000,23.100,0.0000,0.0000,-170.0000
C01265=23.000,-35.000,23.100,0.0000,0.0000,-170.0000
C01266=18.000,-35.000,23.100,0.0000,0.0000,-170.0000
C01267=13.000,-35.000,23.100,0.0000,0.0000,-170.0000
C01268=8.000,-35.000,23.100,0.0000,0.0000,-170.0000
C01269=3.000,-35.000,23.100,0.0000,0.0000,-170.0000
C01270=-2.000,-35.000,23.100,0.0000,0.0000,-170.0000
C01271=-7.000,-35.000,23.100,0.0000,0.0000,-170.0000
C01272=-12.000,-35.000,23.100,0.0000,0.0000,-170.0000
C01273=-17.000,-35.000,23.100,0.0000,0.0000,-170.0000
C01274=-22.000,-35.000,23.100,0.0000,0.0000,-170.0000
C01275=-27.000,-35.000,23.100,0.0000,0.0000,-170.0000
C01276=-27.000,-35.000,24.800,0.0000,0.0000,-170.0000
C01277=-22.000,-35.000,24.800,0.0000,0.0000,-170.0000
C01278=-17.000,-35.000,24.800,0.0000,0.0000,-170.0000
C01279=-12.000,-35.000,24.800,0.0000,0.0000,-170.0000
C01280=-7.000,-35.000,24.800,0.0000,0.0000,-170.0000
C01281=-2.000,-35.000,24.800,0.0000,0.0000,-170.0000
C01282=3.000,-35.000,24.800,0.0000,0.0000,-170.0000
C01283=8.000,-35.000,24.800,0.0000,0.0000,-170.0000
C01284=13.000,-35.000,24.800,0.0000,0.0000,-170.0000
C01285=18.000,-35.000,24.800,0.0000,0.0000,-170.0000
C01286=23.000,-35.000,24.800,0.0000,0.0000,-170.0000
C01287=28.000,-35.000,24.800,0.0000,0.0000,-170.0000
C01288=33.000,-35.000,24.800,0.0000,0.0000,-170.0000
C01289=38.000,-35.000,24.800,0.0000,0.0000,-170.0000
C01290=43.000,-35.000,24.800,0.0000,0.0000,-170.0000
C01291=48.000,-35.000,24.800,0.0000,0.0000,-170.0000
C01292=53.000,-35.000,24.800,0.0000,0.0000,-170.0000
C01293=58.000,-35.000,24.800,0.0000,0.0000,-170.0000
C01294=63.000,-35.000,24.800,0.0000,0.0000,-170.0000
C01295=68.000,-35.000,24.800,0.0000,0.0000,-170.0000
C01296=73.000,-35.000,24.800,0.0000,0.0000,-170.0000
C01297=73.000,-35.000,24.800,0.0000,0.0000,-170.0000
C01298=75.750,-32.250,24.800,0.0000,0.0000,-170.0000
C01299=73.000,-29.500,24.800,0.0000,0.0000,-170.0000
C01300=68.275,-29.500,24.800,0.0000,0.0000,-170.0000
C01301=63.550,-29.500,24.800,0.0000,0.0000,-170.0000
C01302=58.825,-29.500,24.800,0.0000,0.0000,-170.0000
C01303=54.100,-29.500,24.800,0.0000,0.0000,-170.0000
C01304=49.375,-29.500,24.800,0.0000,0.0000,-170.0000
C01305=44.650,-29.500,24.800,0.0000,0.0000,-170.0000
C01306=39.925,-29.500,24.800,0.0000,0.0000,-170.0000
C01307=35.200,-29.500,24.800,0.0000,0.0000,-170.0000
C01308=30.475,-29.500,24.800,0.0000,0.0000,-170.0000
C01309=25.750,-29.500,24.800,0.0000,0.0000,-170.0000
C01310=25.750,-24.500,24.800,0.0000,0.0000,-170.0000
C01311=25.750,-19.500,24.800,0.0000,0.0000,-170.0000
C01312=25.750,-14.500,24.800,0.0000,0.0000,-170.0000
C01313=25.750,-9.500,24.800,0.0000,0.0000,-170.0000
C01314=25.750,-4.500,24.800,0.0000,0.0000,-170.0000
C01315=25.750,0.500,24.800,0.0000,0.0000,-170.0000
C01316=25.750,5.500,24.800,0.0000,0.0000,-170.0000
C01317=25.750,10.500,24.800,0.0000,0.0000,-170.0000
C01318=25.750,15.500,24.800,0.0000,0.0000,-170.0000
C01319=25.750,20.500,24.800,0.0000,0.0000,-170.0000
C01320=25.750,25.500,24.800,0.0000,0.0000,-170.0000
C01321=25.750,30.500,24.800,0.0000,0.0000,-170.0000
C01322=25.750,35.500,24.800,0.0000,0.0000,-170.0000
C01323=25.750,40.500,24.800,0.0000,0.0000,-170.0000
C01324=25.750,45.500,24.800,0.0000,0.0000,-170.0000
C01325=25.750,50.500,24.800,0.0000,0.0000,-170.0000
C01326=25.750,55.500,24.800,0.0000,0.0000,-170.0000
C01327=25.750,60.500,24.800,0.0000,0.0000,-170.0000
C01328=25.750,65.500,24.800,0.0000,0.0000,-170.0000
C01329=25.750,70.500,24.800,0.0000,0.0000,-170.0000
C01330=25.750,75.500,24.800,0.0000,0.0000,-170.0000
C01331=25.750,80.500,24.800,0.0000,0.0000,-170.0000
C01332=25.750,80.500,24.800,0.0000,0.0000,-170.0000
C01333=23.000,83.250,24.800,0.0000,0.0000,-170.0000
C01334=20.250,80.500,24.800,0.0000,0.0000,-170.0000
C01335=20.250,75.500,24.800,0.0000,0.0000,-170.0000
C01336=20.250,70.500,24.800,0.0000,0.0000,-170.0000
C01337=20.250,65.500,24.800,0.0000,0.0000,-170.0000
C01338=20.250,60.500,24.800,0.0000,0.0000,-170.0000
C01339=20.250,55.500,24.800,0.0000,0.0000,-170.0000
C01340=20.250,50.500,24.800,0.0000,0.0000,-170.0000
C01341=20.250,45.500,24.800,0.0000,0.0000,-170.0000
C01342=20.250,40.500,24.800,0.0000,0.0000,-170.0000
C01343=20.250,35.500,24.800,0.0000,0.0000,-170.0000
C01344=20.250,30.500,24.800,0.0000,0.0000,-170.0000
C01345=20.250,25.500,24.800,0.0000,0.0000,-170.0000
C01346=20.250,20.500,24.800,0.0000,0.0000,-170.0000
C01347=20.250,15.500,24.800,0.0000,0.0000,-170.0000
C01348=20.250,10.500,24.800,0.0000,0.0000,-170.0000
C01349=20.250,5.500,24.800,0.0000,0.0000,-170.0000
C01350=20.250,0.500,24.800,0.0000,0.0000,-170.0000
C01351=20.250,-4.500,24.800,0.0000,0.0000,-170.0000
C01352=20.250,-9.500,24.800,0.0000,0.0000,-170.0000
C01353=20.250,-14.500,24.800,0.0000,0.0000,-170.0000
C01354=20.250,-19.500,24.800,0.0000,0.0000,-170.0000
C01355=20.250,-24.500,24.800,0.0000,0.0000,-170.0000
C01356=20.250,-29.500,24.800,0.0000,0.0000,-170.0000
C01357=15.525,-29.500,24.800,0.0000,0.0000,-170.0000
C01358=10.800,-29.500,24.800,0.0000,0.0000,-170.0000
C01359=6.075,-29.500,24.800,0.0000,0.0000,-170.0000
C01360=1.350,-29.500,24.800,0.0000,0.0000,-170.0000
C01361=-3.375,-29.500,24.800,0.0000,0.0000,-170.0000
C01362=-8.100,-29.500,24.800,0.0000,0.0000,-170.0000
C01363=-12.825,-29.500,24.800,0.0000,0.0000,-170.0000
C01364=-17.550,-29.500,24.800,0.0000,0.0000,-170.0000
C01365=-22.275,-29.500,24.800,0.0000,0.0000,-170.0000
C01366=-27.000,-29.500,24.800,0.0000,0.0000,-170.0000
C01367=-27.000,-29.500,150.000,0.0000,0.0000,-170.0000
C01368=185.000,150.000,150.000,0.0000,0.0000,-170.0000
//INST
///DATE 2026/11/04 18:55
///ATTR SC,RW,RJ
////FRAME USER 9
///GROUP1 RB1
NOP
MOVJ C00000 VJ=0.78
MOVJ C00001 VJ=0.78
MOVL C00002 V=11.0 ACC=20 DEC=20
*LAG1
MACRO1 MJ#(0) ARGF1
ARCON
MOVL C00003 V=7.0 ACC=20 DEC=20
MOVL C00004 V=7.0 ACC=20 DEC=20
MOVL C00005 V=7.0 ACC=20 DEC=20
MOVL C00006 V=7.0 ACC=20 DEC=20
MOVL C00007 V=7.0 ACC=20 DEC=20
MOVL C00008 V=7.0 ACC=20 DEC=20
MOVL C00009 V=7.0 ACC=20 DEC=20
MOVL C00010 V=7.0 ACC=20 DEC=20
MOVL C00011 V=7.0 ACC=20 DEC=20
MOVL C00012 V=7.0 ACC=20 DEC=20
MOVL C00013 V=7.0 ACC=20 DEC=20
MOVL C00014 V=7.0 ACC=20 DEC=20
MOVL C00015 V=7.0 ACC=20 DEC=20
MOVL C00016 V=7.0 ACC=20 DEC=20
MOVL C00017 V=7.0 ACC=20 DEC=20
MOVL C00018 V=7.0 ACC=20 DEC=20
MOVL C00019 V=7.0 ACC=20 DEC=20
MOVL C00020 V=7.0 ACC=20 DEC=20
MOVL C00021 V=7.0 ACC=20 DEC=20
MOVL C00022 V=11.0 ACC=20 DEC=20
MOVC C00023 V=11.0 ACC=20 DEC=20
MOVC C00024 V=11.0 ACC=20 DEC=20
MOVC C00025 V=11.0 ACC=20 DEC=20
MOVL C00026 V=7.0 ACC=20 DEC=20
MOVL C00027 V=7.0 ACC=20 DEC=20
MOVL C00028 V=7.0 ACC=20 DEC=20
MOVL C00029 V=7.0 ACC=20 DEC=20
MOVL C00030 V=7.0 ACC=20 DEC=20
MOVL C00031 V=7.0 ACC=20 DEC=20
MOVL C00032 V=7.0 ACC=20 DEC=20
MOVL C00033 V=7.0 ACC=20 DEC=20
MOVL C00034 V=7.0 ACC=20 DEC=20
MOVL C00035 V=7.0 PL=1
MOVL C00036 V=7.0 ACC=20 DEC=20
MOVL C00037 V=7.0 ACC=20 DEC=20
MOVL C00038 V=7.0 ACC=20 DEC=20
MOVL C00039 V=7.0 ACC=20 DEC=20
MOVL C00040 V=7.0 ACC=20 DEC=20
MOVL C00041 V=7.0 ACC=20 DEC=20
MOVL C00042 V=7.0 ACC=20 DEC=20
MOVL C00043 V=7.0 ACC=20 DEC=20
MOVL C00044 V=7.0 ACC=20 DEC=20
MOVL C00045 V=7.0 ACC=20 DEC=20
MOVL C00046 V=7.0 ACC=20 DEC=20
MOVL C00047 V=7.0 ACC=20 DEC=20
MOVL C00048 V=7.0 ACC=20 DEC=20
MOVL C00049 V=7.0 ACC=20 DEC=20
MOVL C00050 V=7.0 ACC=20 DEC=20
MOVL C00051 V=7.0 ACC=20 DEC=20
MOVL C00052 V=7.0 ACC=20 DEC=20
MOVL C00053 V=7.0 ACC=20 DEC=20
MOVL C00054 V=7.0 ACC=20 DEC=20
MOVL C00055 V=7.0 ACC=20 DEC=20
MOVL C00056 V=7.0 ACC=20 DEC=20
MOVL C00057 V=11.0 ACC=20 DEC=20
MOVC C00058 V=11.0 ACC=20 DEC=20
MOVC C00059 V=11.0 ACC=20 DEC=20
MOVC C00060 V=11.0 ACC=20 DEC=20
MOVL C00061 V=7.0 ACC=20 DEC=20
MOVL C00062 V=7.0 ACC=20 DEC=20
MOVL C00063 V=7.0 ACC=20 DEC=20
MOVL C00064 V=7.0 ACC=20 DEC=20
MOVL C00065 V=7.0 ACC=20 DEC=20
MOVL C00066 V=7.0 ACC=20 DEC=20
MOVL C00067 V=7.0 ACC=20 DEC=20
MOVL C00068 V=7.0 ACC=20 DEC=20
MOVL C00069 V=7.0 ACC=20 DEC=20
MOVL C00070 V=7.0 ACC=20 DEC=20
MOVL C00071 V=7.0 ACC=20 DEC=20
MOVL C00072 V=7.0 ACC=20 DEC=20
MOVL C00073 V=7.0 ACC=20 DEC=20
MOVL C00074 V=7.0 ACC=20 DEC=20
MOVL C00075 V=7.0 ACC=20 DEC=20
MOVL C00076 V=7.0 ACC=20 DEC=20
MOVL C00077 V=7.0 ACC=20 DEC=20
MOVL C00078 V=7.0 ACC=20 DEC=20
MOVL C00079 V=7.0 ACC=20 DEC=20
MOVL C00080 V=7.0 ACC=20 DEC=20
MOVL C00081 V=7.0 ACC=20 DEC=20
MOVL C00082 V=7.0 PL=1
MOVL C00083 V=7.0 ACC=20 DEC=20
MOVL C00084 V=7.0 ACC=20 DEC=20
MOVL C00085 V=7.0 ACC=20 DEC=20
MOVL C00086 V=7.0 ACC=20 DEC=20
MOVL C00087 V=7.0 ACC=20 DEC=20
MOVL C00088 V=7.0 ACC=20 DEC=20
MOVL C00089 V=7.0 ACC=20 DEC=20
MOVL C00090 V=7.0 ACC=20 DEC=20
MOVL C00091 V=7.0 ACC=20 DEC=20
MOVL C00092 V=7.0 ACC=20 DEC=20
ARCOF
TIMER T=30
MOVL C00093 V=11.0 ACC=20 DEC=20
*LAG2
MACRO1 MJ#(0) ARGF2
ARCON
MOVL C00094 V=7.0 ACC=20 DEC=20
MOVL C00095 V=7.0 ACC=20 DEC=20
MOVL C00096 V=7.0 ACC=20 DEC=20
MOVL C00097 V=7.0 ACC=20 DEC=20
MOVL C00098 V=7.0 ACC=20 DEC=20
MOVL C00099 V=7.0 ACC=20 DEC=20
MOVL C00100 V=7.0 ACC=20 DEC=20
MOVL C00101 V=7.0 ACC=20 DEC=20
MOVL C00102 V=7.0 ACC=20 DEC=20
MOVL C00103 V=7.0 PL=1
MOVL C00104 V=7.0 ACC=20 DEC=20
MOVL C00105 V=7.0 ACC=20 DEC=20
MOVL C00106 V=7.0 ACC=20 DEC=20
MOVL C00107 V=7.0 ACC=20 DEC=20
MOVL C00108 V=7.0 ACC=20 DEC=20
MOVL C00109 V=7.0 ACC=20 DEC=20
MOVL C00110 V=7.0 ACC=20 DEC=20
MOVL C00111 V=7.0 ACC=20 DEC=20
MOVL C00112 V=7.0 ACC=20 DEC=20
MOVL C00113 V=7.0 ACC=20 DEC=20
MOVL C00114 V=7.0 ACC=20 DEC=20
MOVL C00115 V=7.0 ACC=20 DEC=20
MOVL C00116 V=7.0 ACC=20 DEC=20
MOVL C00117 V=7.0 ACC=20 DEC=20
MOVL C00118 V=7.0 ACC=20 DEC=20
MOVL C00119 V=7.0 ACC=20 DEC=20
MOVL C00120 V=7.0 ACC=20 DEC=20
MOVL C00121 V=7.0 ACC=20 DEC=20
MOVL C00122 V=7.0 ACC=20 DEC=20
MOVL C00123 V=7.0 ACC=20 DEC=20
MOVL C00124 V=7.0 ACC=20 DEC=20
MOVL C00125 V=11.0 ACC=20 DEC=20
MOVC C00126 V=11.0 ACC=20 DEC=20
MOVC C00127 V=11.0 ACC=20 DEC=20
MOVC C00128 V=11.0 ACC=20 DEC=20
MOVL C00129 V=7.0 ACC=20 DEC=20
MOVL C00130 V=7.0 ACC=20 DEC=20
MOVL C00131 V=7.0 ACC=20 DEC=20
MOVL C00132 V=7.0 ACC=20 DEC=20
MOVL C00133 V=7.0 ACC=20 DEC=20
MOVL C00134 V=7.0 ACC=20 DEC=20
MOVL C00135 V=7.0 ACC=20 DEC=20
MOVL C00136 V=7.0 ACC=20 DEC=20
MOVL C00137 V=7.0 ACC=20 DEC=20
MOVL C00138 V=7.0 ACC=20 DEC=20
MOVL C00139 V=7.0 ACC=20 DEC=20
MOVL C00140 V=7.0 ACC=20 DEC=20
MOVL C00141 V=7.0 ACC=20 DEC=20
MOVL C00142 V=7.0 ACC=20 DEC=20
MOVL C00143 V=7.0 ACC=20 DEC=20
MOVL C00144 V=7.0 ACC=20 DEC=20
MOVL C00145 V=7.0 ACC=20 DEC=20
MOVL C00146 V=7.0 ACC=20 DEC=20
MOVL C00147 V=7.0 ACC=20 DEC=20
MOVL C00148 V=7.0 ACC=20 DEC=20
MOVL C00149 V=7.0 ACC=20 DEC=20
MOVL C00150 V=7.0 PL=1
MOVL C00151 V=7.0 ACC=20 DEC=20
MOVL C00152 V=7.0 ACC=20 DEC=20
MOVL C00153 V=7.0 ACC=20 DEC=20
MOVL C00154 V=7.0 ACC=20 DEC=20
MOVL C00155 V=7.0 ACC=20 DEC=20
MOVL C00156 V=7.0 ACC=20 DEC=20
MOVL C00157 V=7.0 ACC=20 DEC=20
MOVL C00158 V=7.0 ACC=20 DEC=20
MOVL C00159 V=7.0 ACC=20 DEC=20
MOVL C00160 V=11.0 ACC=20 DEC=20
MOVC C00161 V=11.0 ACC=20 DEC=20
MOVC C00162 V=11.0 ACC=20 DEC=20
MOVC C00163 V=11.0 ACC=20 DEC=20
MOVL C00164 V=7.0 ACC=20 DEC=20
MOVL C00165 V=7.0 ACC=20 DEC=20
MOVL C00166 V=7.0 ACC=20 DEC=20
MOVL C00167 V=7.0 ACC=20 DEC=20
MOVL C00168 V=7.0 ACC=20 DEC=20
MOVL C00169 V=7.0 ACC=20 DEC=20
MOVL C00170 V=7.0 ACC=20 DEC=20
MOVL C00171 V=7.0 ACC=20 DEC=20
MOVL C00172 V=7.0 ACC=20 DEC=20
MOVL C00173 V=7.0 ACC=20 DEC=20
MOVL C00174 V=7.0 ACC=20 DEC=20
MOVL C00175 V=7.0 ACC=20 DEC=20
MOVL C00176 V=7.0 ACC=20 DEC=20
MOVL C00177 V=7.0 ACC=20 DEC=20
MOVL C00178 V=7.0 ACC=20 DEC=20
MOVL C00179 V=7.0 ACC=20 DEC=20
MOVL C00180 V=7.0 ACC=20 DEC=20
MOVL C00181 V=7.0 ACC=20 DEC=20
MOVL C00182 V=7.0 ACC=20 DEC=20
MOVL C00183 V=7.0 ACC=20 DEC=20
ARCOF
TIMER T=30
MOVL C00184 V=11.0 ACC=20 DEC=20
*LAG3
MACRO1 MJ#(0) ARGF2
ARCON
MOVL C00185 V=7.0 ACC=20 DEC=20
MOVL C00186 V=7.0 ACC=20 DEC=20
MOVL C00187 V=7.0 ACC=20 DEC=20
MOVL C00188 V=7.0 ACC=20 DEC=20
MOVL C00189 V=7.0 ACC=20 DEC=20
MOVL C00190 V=7.0 ACC=20 DEC=20
MOVL C00191 V=7.0 ACC=20 DEC=20
MOVL C00192 V=7.0 ACC=20 DEC=20
MOVL C00193 V=7.0 ACC=20 DEC=20
MOVL C00194 V=7.0 ACC=20 DEC=20
MOVL C00195 V=7.0 ACC=20 DEC=20
MOVL C00196 V=7.0 ACC=20 DEC=20
MOVL C00197 V=7.0 ACC=20 DEC=20
MOVL C00198 V=7.0 ACC=20 DEC=20
MOVL C00199 V=7.0 ACC=20 DEC=20
MOVL C00200 V=7.0 ACC=20 DEC=20
MOVL C00201 V=7.0 ACC=20 DEC=20
MOVL C00202 V=7.0 ACC=20 DEC=20
MOVL C00203 V=7.0 ACC=20 DEC=20
MOVL C00204 V=11.0 ACC=20 DEC=20
MOVC C00205 V=11.0 ACC=20 DEC=20
MOVC C00206 V=11.0 ACC=20 DEC=20
MOVC C00207 V=11.0 ACC=20 DEC=20
MOVL C00208 V=7.0 ACC=20 DEC=20
MOVL C00209 V=7.0 ACC=20 DEC=20
MOVL C00210 V=7.0 ACC=20 DEC=20
MOVL C00211 V=7.0 ACC=20 DEC=20
MOVL C00212 V=7.0 ACC=20 DEC=20
MOVL C00213 V=7.0 ACC=20 DEC=20
MOVL C00214 V=7.0 ACC=20 DEC=20
MOVL C00215 V=7.0 ACC=20 DEC=20
MOVL C00216 V=7.0 ACC=20 DEC=20
MOVL C00217 V=7.0 PL=1
MOVL C00218 V=7.0 ACC=20 DEC=20
MOVL C00219 V=7.0 ACC=20 DEC=20
MOVL C00220 V=7.0 ACC=20 DEC=20
MOVL C00221 V=7.0 ACC=20 DEC=20
MOVL C00222 V=7.0 ACC=20 DEC=20
MOVL C00223 V=7.0 ACC=20 DEC=20
MOVL C00224 V=7.0 ACC=20 DEC=20
MOVL C00225 V=7.0 ACC=20 DEC=20
MOVL C00226 V=7.0 ACC=20 DEC=20
MOVL C00227 V=7.0 ACC=20 DEC=20
MOVL C00228 V=7.0 ACC=20 DEC=20
MOVL C00229 V=7.0 ACC=20 DEC=20
MOVL C00230 V=7.0 ACC=20 DEC=20
MOVL C00231 V=7.0 ACC=20 DEC=20
MOVL C00232 V=7.0 ACC=20 DEC=20
MOVL C00233 V=7.0 ACC=20 DEC=20
MOVL C00234 V=7.0 ACC=20 DEC=20
MOVL C00235 V=7.0 ACC=20 DEC=20
MOVL C00236 V=7.0 ACC=20 DEC=20
MOVL C00237 V=7.0 ACC=20 DEC=20
MOVL C00238 V=7.0 ACC=20 DEC=20
MOVL C00239 V=11.0 ACC=20 DEC=20
MOVC C00240 V=11.0 ACC=20 DEC=20
MOVC C00241 V=11.0 ACC=20 DEC=20
MOVC C00242 V=11.0 ACC=20 DEC=20
MOVL C00243 V=7.0 ACC=20 DEC=20
MOVL C00244 V=7.0 ACC=20 DEC=20
MOVL C00245 V=7.0 ACC=20 DEC=20
MOVL C00246 V=7.0 ACC=20 DEC=20
MOVL C00247 V=7.0 ACC=20 DEC=20
MOVL C00248 V=7.0 ACC=20 DEC=20
MOVL C00249 V=7.0 ACC=20 DEC=20
MOVL C00250 V=7.0 ACC=20 DEC=20
MOVL C00251 V=7.0 ACC=20 DEC=20
MOVL C00252 V=7.0 ACC=20 DEC=20
MOVL C00253 V=7.0 ACC=20 DEC=20
MOVL C00254 V=7.0 ACC=20 DEC=20
MOVL C00255 V=7.0 ACC=20 DEC=20
MOVL C00256 V=7.0 ACC=20 DEC=20
MOVL C00257 V=7.0 ACC=20 DEC=20
MOVL C00258 V=7.0 ACC=20 DEC=20
MOVL C00259 V=7.0 ACC=20 DEC=20
MOVL C00260 V=7.0 ACC=20 DEC=20
MOVL C00261 V=7.0 ACC=20 DEC=20
MOVL C00262 V=7.0 ACC=20 DEC=20
MOVL C00263 V=7.0 ACC=20 DEC=20
MOVL C00264 V=7.0 PL=1
MOVL C00265 V=7.0 ACC=20 DEC=20
MOVL C00266 V=7.0 ACC=20 DEC=20
MOVL C00267 V=7.0 ACC=20 DEC=20
MOVL C00268 V=7.0 ACC=20 DEC=20
MOVL C00269 V=7.0 ACC=20 DEC=20
MOVL C00270 V=7.0 ACC=20 DEC=20
MOVL C00271 V=7.0 ACC=20 DEC=20
MOVL C00272 V=7.0 ACC=20 DEC=20
MOVL C00273 V=7.0 ACC=20 DEC=20
MOVL C00274 V=7.0 ACC=20 DEC=20
ARCOF
TIMER T=30
MOVL C00275 V=11.0 ACC=20 DEC=20
*LAG4
MACRO1 MJ#(0) ARGF2
ARCON
MOVL C00276 V=7.0 ACC=20 DEC=20
MOVL C00277 V=7.0 ACC=20 DEC=20
MOVL C00278 V=7.0 ACC=20 DEC=20
MOVL C00279 V=7.0 ACC=20 DEC=20
MOVL C00280 V=7.0 ACC=20 DEC=20
MOVL C00281 V=7.0 ACC=20 DEC=20
MOVL C00282 V=7.0 ACC=20 DEC=20
MOVL C00283 V=7.0 ACC=20 DEC=20
MOVL C00284 V=7.0 ACC=20 DEC=20
MOVL C00285 V=7.0 PL=1
MOVL C00286 V=7.0 ACC=20 DEC=20
MOVL C00287 V=7.0 ACC=20 DEC=20
MOVL C00288 V=7.0 ACC=20 DEC=20
MOVL C00289 V=7.0 ACC=20 DEC=20
MOVL C00290 V=7.0 ACC=20 DEC=20
MOVL C00291 V=7.0 ACC=20 DEC=20
MOVL C00292 V=7.0 ACC=20 DEC=20
MOVL C00293 V=7.0 ACC=20 DEC=20
MOVL C00294 V=7.0 ACC=20 DEC=20
MOVL C00295 V=7.0 ACC=20 DEC=20
MOVL C00296 V=7.0 ACC=20 DEC=20
MOVL C00297 V=7.0 ACC=20 DEC=20
MOVL C00298 V=7.0 ACC=20 DEC=20
MOVL C00299 V=7.0 ACC=20 DEC=20
MOVL C00300 V=7.0 ACC=20 DEC=20
MOVL C00301 V=7.0 ACC=20 DEC=20
MOVL C00302 V=7.0 ACC=20 DEC=20
MOVL C00303 V=7.0 ACC=20 DEC=20
MOVL C00304 V=7.0 ACC=20 DEC=20
MOVL C00305 V=7.0 ACC=20 DEC=20
MOVL C00306 V=7.0 ACC=20 DEC=20
MOVL C00307 V=11.0 ACC=20 DEC=20
MOVC C00308 V=11.0 ACC=20 DEC=20
MOVC C00309 V=11.0 ACC=20 DEC=20
MOVC C00310 V=11.0 ACC=20 DEC=20
MOVL C00311 V=7.0 ACC=20 DEC=20
MOVL C00312 V=7.0 ACC=20 DEC=20
MOVL C00313 V=7.0 ACC=20 DEC=20
MOVL C00314 V=7.0 ACC=20 DEC=20
MOVL C00315 V=7.0 ACC=20 DEC=20
MOVL C00316 V=7.0 ACC=20 DEC=20
MOVL C00317 V=7.0 ACC=20 DEC=20
MOVL C00318 V=7.0 ACC=20 DEC=20
MOVL C00319 V=7.0 ACC=20 DEC=20
MOVL C00320 V=7.0 ACC=20 DEC=20
MOVL C00321 V=7.0 ACC=20 DEC=20
MOVL C00322 V=7.0 ACC=20 DEC=20
MOVL C00323 V=7.0 ACC=20 DEC=20
MOVL C00324 V=7.0 ACC=20 DEC=20
MOVL C00325 V=7.0 ACC=20 DEC=20
MOVL C00326 V=7.0 ACC=20 DEC=20
MOVL C00327 V=7.0 ACC=20 DEC=20
MOVL C00328 V=7.0 ACC=20 DEC=20
MOVL C00329 V=7.0 ACC=20 DEC=20
MOVL C00330 V=7.0 ACC=20 DEC=20
MOVL C00331 V=7.0 ACC=20 DEC=20
MOVL C00332 V=7.0 PL=1
MOVL C00333 V=7.0 ACC=20 DEC=20
MOVL C00334 V=7.0 ACC=20 DEC=20
MOVL C00335 V=7.0 ACC=20 DEC=20
MOVL C00336 V=7.0 ACC=20 DEC=20
MOVL C00337 V=7.0 ACC=20 DEC=20
MOVL C00338 V=7.0 ACC=20 DEC=20
MOVL C00339 V=7.0 ACC=20 DEC=20
MOVL C00340 V=7.0 ACC=20 DEC=20
MOVL C00341 V=7.0 ACC=20 DEC=20
MOVL C00342 V=11.0 ACC=20 DEC=20
MOVC C00343 V=11.0 ACC=20 DEC=20
MOVC C00344 V=11.0 ACC=20 DEC=20
MOVC C00345 V=11.0 ACC=20 DEC=20
MOVL C00346 V=7.0 ACC=20 DEC=20
MOVL C00347 V=7.0 ACC=20 DEC=20
MOVL C00348 V=7.0 ACC=20 DEC=20
MOVL C00349 V=7.0 ACC=20 DEC=20
MOVL C00350 V=7.0 ACC=20 DEC=20
MOVL C00351 V=7.0 ACC=20 DEC=20
MOVL C00352 V=7.0 ACC=20 DEC=20
MOVL C00353 V=7.0 ACC=20 DEC=20
MOVL C00354 V=7.0 ACC=20 DEC=20
MOVL C00355 V=7.0 ACC=20 DEC=20
MOVL C00356 V=7.0 ACC=20 DEC=20
MOVL C00357 V=7.0 ACC=20 DEC=20
MOVL C00358 V=7.0 ACC=20 DEC=20
MOVL C00359 V=7.0 ACC=20 DEC=20
MOVL C00360 V=7.0 ACC=20 DEC=20
MOVL C00361 V=7.0 ACC=20 DEC=20
MOVL C00362 V=7.0 ACC=20 DEC=20
MOVL C00363 V=7.0 ACC=20 DEC=20
MOVL C00364 V=7.0 ACC=20 DEC=20
MOVL C00365 V=7.0 ACC=20 DEC=20
ARCOF
TIMER T=30
MOVL C00366 V=11.0 ACC=20 DEC=20
*LAG5
MACRO1 MJ#(0) ARGF2
ARCON
MOVL C00367 V=7.0 ACC=20 DEC=20
MOVL C00368 V=7.0 ACC=20 DEC=20
MOVL C00369 V=7.0 ACC=20 DEC=20
MOVL C00370 V=7.0 ACC=20 DEC=20
MOVL C00371 V=7.0 ACC=20 DEC=20
MOVL C00372 V=7.0 ACC=20 DEC=20
MOVL C00373 V=7.0 ACC=20 DEC=20
MOVL C00374 V=7.0 ACC=20 DEC=20
MOVL C00375 V=7.0 ACC=20 DEC=20
MOVL C00376 V=7.0 ACC=20 DEC=20
MOVL C00377 V=7.0 ACC=20 DEC=20
MOVL C00378 V=7.0 ACC=20 DEC=20
MOVL C00379 V=7.0 ACC=20 DEC=20
MOVL C00380 V=7.0 ACC=20 DEC=20
MOVL C00381 V=7.0 ACC=20 DEC=20
MOVL C00382 V=7.0 ACC=20 DEC=20
MOVL C00383 V=7.0 ACC=20 DEC=20
MOVL C00384 V=7.0 ACC=20 DEC=20
MOVL C00385 V=7.0 ACC=20 DEC=20
MOVL C00386 V=11.0 ACC=20 DEC=20
MOVC C00387 V=11.0 ACC=20 DEC=20
MOVC C00388 V=11.0 ACC=20 DEC=20
MOVC C00389 V=11.0 ACC=20 DEC=20
MOVL C00390 V=7.0 ACC=20 DEC=20
MOVL C00391 V=7.0 ACC=20 DEC=20
MOVL C00392 V=7.0 ACC=20 DEC=20
MOVL C00393 V=7.0 ACC=20 DEC=20
MOVL C00394 V=7.0 ACC=20 DEC=20
MOVL C00395 V=7.0 ACC=20 DEC=20
MOVL C00396 V=7.0 ACC=20 DEC=20
MOVL C00397 V=7.0 ACC=20 DEC=20
MOVL C00398 V=7.0 ACC=20 DEC=20
MOVL C00399 V=7.0 PL=1
MOVL C00400 V=7.0 ACC=20 DEC=20
MOVL C00401 V=7.0 ACC=20 DEC=20
MOVL C00402 V=7.0 ACC=20 DEC=20
MOVL C00403 V=7.0 ACC=20 DEC=20
MOVL C00404 V=7.0 ACC=20 DEC=20
MOVL C00405 V=7.0 ACC=20 DEC=20
MOVL C00406 V=7.0 ACC=20 DEC=20
MOVL C00407 V=7.0 ACC=20 DEC=20
MOVL C00408 V=7.0 ACC=20 DEC=20
MOVL C00409 V=7.0 ACC=20 DEC=20
MOVL C00410 V=7.0 ACC=20 DEC=20
MOVL C00411 V=7.0 ACC=20 DEC=20
MOVL C00412 V=7.0 ACC=20 DEC=20
MOVL C00413 V=7.0 ACC=20 DEC=20
MOVL C00414 V=7.0 ACC=20 DEC=20
MOVL C00415 V=7.0 ACC=20 DEC=20
MOVL C00416 V=7.0 ACC=20 DEC=20
MOVL C00417 V=7.0 ACC=20 DEC=20
MOVL C00418 V=7.0 ACC=20 DEC=20
MOVL C00419 V=7.0 ACC=20 DEC=20
MOVL C00420 V=7.0 ACC=20 DEC=20
MOVL C00421 V=11.0 ACC=20 DEC=20
MOVC C00422 V=11.0 ACC=20 DEC=20
MOVC C00423 V=11.0 ACC=20 DEC=20
MOVC C00424 V=11.0 ACC=20 DEC=20
MOVL C00425 V=7.0 ACC=20 DEC=20
MOVL C00426 V=7.0 ACC=20 DEC=20
MOVL C00427 V=7.0 ACC=20 DEC=20
MOVL C00428 V=7.0 ACC=20 DEC=20
MOVL C00429 V=7.0 ACC=20 DEC=20
MOVL C00430 V=7.0 ACC=20 DEC=20
MOVL C00431 V=7.0 ACC=20 DEC=20
MOVL C00432 V=7.0 ACC=20 DEC=20
MOVL C00433 V=7.0 ACC=20 DEC=20
MOVL C00434 V=7.0 ACC=20 DEC=20
MOVL C00435 V=7.0 ACC=20 DEC=20
MOVL C00436 V=7.0 ACC=20 DEC=20
MOVL C00437 V=7.0 ACC=20 DEC=20
MOVL C00438 V=7.0 ACC=20 DEC=20
MOVL C00439 V=7.0 ACC=20 DEC=20
MOVL C00440 V=7.0 ACC=20 DEC=20
MOVL C00441 V=7.0 ACC=20 DEC=20
MOVL C00442 V=7.0 ACC=20 DEC=20
MOVL C00443 V=7.0 ACC=20 DEC=20
MOVL C00444 V=7.0 ACC=20 DEC=20
MOVL C00445 V=7.0 ACC=20 DEC=20
MOVL C00446 V=7.0 PL=1
MOVL C00447 V=7.0 ACC=20 DEC=20
MOVL C00448 V=7.0 ACC=20 DEC=20
MOVL C00449 V=7.0 ACC=20 DEC=20
MOVL C00450 V=7.0 ACC=20 DEC=20
MOVL C00451 V=7.0 ACC=20 DEC=20
MOVL C00452 V=7.0 ACC=20 DEC=20
MOVL C00453 V=7.0 ACC=20 DEC=20
MOVL C00454 V=7.0 ACC=20 DEC=20
MOVL C00455 V=7.0 ACC=20 DEC=20
MOVL C00456 V=7.0 ACC=20 DEC=20
ARCOF
TIMER T=30
MOVL C00457 V=11.0 ACC=20 DEC=20
*LAG6
MACRO1 MJ#(0) ARGF2
ARCON
MOVL C00458 V=7.0 ACC=20 DEC=20
MOVL C00459 V=7.0 ACC=20 DEC=20
MOVL C00460 V=7.0 ACC=20 DEC=20
MOVL C00461 V=7.0 ACC=20 DEC=20
MOVL C00462 V=7.0 ACC=20 DEC=20
MOVL C00463 V=7.0 ACC=20 DEC=20
MOVL C00464 V=7.0 ACC=20 DEC=20
MOVL C00465 V=7.0 ACC=20 DEC=20
MOVL C00466 V=7.0 ACC=20 DEC=20
MOVL C00467 V=7.0 PL=1
MOVL C00468 V=7.0 ACC=20 DEC=20
MOVL C00469 V=7.0 ACC=20 DEC=20
MOVL C00470 V=7.0 ACC=20 DEC=20
MOVL C00471 V=7.0 ACC=20 DEC=20
MOVL C00472 V=7.0 ACC=20 DEC=20
MOVL C00473 V=7.0 ACC=20 DEC=20
MOVL C00474 V=7.0 ACC=20 DEC=20
MOVL C00475 V=7.0 ACC=20 DEC=20
MOVL C00476 V=7.0 ACC=20 DEC=20
MOVL C00477 V=7.0 ACC=20 DEC=20
MOVL C00478 V=7.0 ACC=20 DEC=20
MOVL C00479 V=7.0 ACC=20 DEC=20
MOVL C00480 V=7.0 ACC=20 DEC=20
MOVL C00481 V=7.0 ACC=20 DEC=20
MOVL C00482 V=7.0 ACC=20 DEC=20
MOVL C00483 V=7.0 ACC=20 DEC=20
MOVL C00484 V=7.0 ACC=20 DEC=20
MOVL C00485 V=7.0 ACC=20 DEC=20
MOVL C00486 V=7.0 ACC=20 DEC=20
MOVL C00487 V=7.0 ACC=20 DEC=20
MOVL C00488 V=7.0 ACC=20 DEC=20
MOVL C00489 V=11.0 ACC=20 DEC=20
MOVC C00490 V=11.0 ACC=20 DEC=20
MOVC C00491 V=11.0 ACC=20 DEC=20
MOVC C00492 V=11.0 ACC=20 DEC=20
MOVL C00493 V=7.0 ACC=20 DEC=20
MOVL C00494 V=7.0 ACC=20 DEC=20
MOVL C00495 V=7.0 ACC=20 DEC=20
MOVL C00496 V=7.0 ACC=20 DEC=20
MOVL C00497 V=7.0 ACC=20 DEC=20
MOVL C00498 V=7.0 ACC=20 DEC=20
MOVL C00499 V=7.0 ACC=20 DEC=20
MOVL C00500 V=7.0 ACC=20 DEC=20
MOVL C00501 V=7.0 ACC=20 DEC=20
MOVL C00502 V=7.0 ACC=20 DEC=20
MOVL C00503 V=7.0 ACC=20 DEC=20
MOVL C00504 V=7.0 ACC=20 DEC=20
MOVL C00505 V=7.0 ACC=20 DEC=20
MOVL C00506 V=7.0 ACC=20 DEC=20
MOVL C00507 V=7.0 ACC=20 DEC=20
MOVL C00508 V=7.0 ACC=20 DEC=20
MOVL C00509 V=7.0 ACC=20 DEC=20
MOVL C00510 V=7.0 ACC=20 DEC=20
MOVL C00511 V=7.0 ACC=20 DEC=20
MOVL C00512 V=7.0 ACC=20 DEC=20
MOVL C00513 V=7.0 ACC=20 DEC=20
MOVL C00514 V=7.0 PL=1
MOVL C00515 V=7.0 ACC=20 DEC=20
MOVL C00516 V=7.0 ACC=20 DEC=20
MOVL C00517 V=7.0 ACC=20 DEC=20
MOVL C00518 V=7.0 ACC=20 DEC=20
MOVL C00519 V=7.0 ACC=20 DEC=20
MOVL C00520 V=7.0 ACC=20 DEC=20
MOVL C00521 V=7.0 ACC=20 DEC=20
MOVL C00522 V=7.0 ACC=20 DEC=20
MOVL C00523 V=7.0 ACC=20 DEC=20
MOVL C00524 V=11.0 ACC=20 DEC=20
MOVC C00525 V=11.0 ACC=20 DEC=20
MOVC C00526 V=11.0 ACC=20 DEC=20
MOVC C00527 V=11.0 ACC=20 DEC=20
MOVL C00528 V=7.0 ACC=20 DEC=20
MOVL C00529 V=7.0 ACC=20 DEC=20
MOVL C00530 V=7.0 ACC=20 DEC=20
MOVL C00531 V=7.0 ACC=20 DEC=20
MOVL C00532 V=7.0 ACC=20 DEC=20
MOVL C00533 V=7.0 ACC=20 DEC=20
MOVL C00534 V=7.0 ACC=20 DEC=20
MOVL C00535 V=7.0 ACC=20 DEC=20
MOVL C00536 V=7.0 ACC=20 DEC=20
MOVL C00537 V=7.0 ACC=20 DEC=20
MOVL C00538 V=7.0 ACC=20 DEC=20
MOVL C00539 V=7.0 ACC=20 DEC=20
MOVL C00540 V=7.0 ACC=20 DEC=20
MOVL C00541 V=7.0 ACC=20 DEC=20
MOVL C00542 V=7.0 ACC=20 DEC=20
MOVL C00543 V=7.0 ACC=20 DEC=20
MOVL C00544 V=7.0 ACC=20 DEC=20
MOVL C00545 V=7.0 ACC=20 DEC=20
MOVL C00546 V=7.0 ACC=20 DEC=20
MOVL C00547 V=7.0 ACC=20 DEC=20
ARCOF
TIMER T=30
MOVL C00548 V=11.0 ACC=20 DEC=20
*LAG7
MACRO1 MJ#(0) ARGF2
ARCON
MOVL C00549 V=7.0 ACC=20 DEC=20
MOVL C00550 V=7.0 ACC=20 DEC=20
MOVL C00551 V=7.0 ACC=20 DEC=20
MOVL C00552 V=7.0 ACC=20 DEC=20
MOVL C00553 V=7.0 ACC=20 DEC=20
MOVL C00554 V=7.0 ACC=20 DEC=20
MOVL C00555 V=7.0 ACC=20 DEC=20
MOVL C00556 V=7.0 ACC=20 DEC=20
MOVL C00557 V=7.0 ACC=20 DEC=20
MOVL C00558 V=7.0 ACC=20 DEC=20
MOVL C00559 V=7.0 ACC=20 DEC=20
MOVL C00560 V=7.0 ACC=20 DEC=20
MOVL C00561 V=7.0 ACC=20 DEC=20
MOVL C00562 V=7.0 ACC=20 DEC=20
MOVL C00563 V=7.0 ACC=20 DEC=20
MOVL C00564 V=7.0 ACC=20 DEC=20
MOVL C00565 V=7.0 ACC=20 DEC=20
MOVL C00566 V=7.0 ACC=20 DEC=20
MOVL C00567 V=7.0 ACC=20 DEC=20
MOVL C00568 V=11.0 ACC=20 DEC=20
MOVC C00569 V=11.0 ACC=20 DEC=20
MOVC C00570 V=11.0 ACC=20 DEC=20
MOVC C00571 V=11.0 ACC=20 DEC=20
MOVL C00572 V=7.0 ACC=20 DEC=20
MOVL C00573 V=7.0 ACC=20 DEC=20
MOVL C00574 V=7.0 ACC=20 DEC=20
MOVL C00575 V=7.0 ACC=20 DEC=20
MOVL C00576 V=7.0 ACC=20 DEC=20
MOVL C00577 V=7.0 ACC=20 DEC=20
MOVL C00578 V=7.0 ACC=20 DEC=20
MOVL C00579 V=7.0 ACC=20 DEC=20
MOVL C00580 V=7.0 ACC=20 DEC=20
MOVL C00581 V=7.0 PL=1
MOVL C00582 V=7.0 ACC=20 DEC=20
MOVL C00583 V=7.0 ACC=20 DEC=20
MOVL C00584 V=7.0 ACC=20 DEC=20
MOVL C00585 V=7.0 ACC=20 DEC=20
MOVL C00586 V=7.0 ACC=20 DEC=20
MOVL C00587 V=7.0 ACC=20 DEC=20
MOVL C00588 V=7.0 ACC=20 DEC=20
MOVL C00589 V=7.0 ACC=20 DEC=20
MOVL C00590 V=7.0 ACC=20 DEC=20
MOVL C00591 V=7.0 ACC=20 DEC=20
MOVL C00592 V=7.0 ACC=20 DEC=20
MOVL C00593 V=7.0 ACC=20 DEC=20
MOVL C00594 V=7.0 ACC=20 DEC=20
MOVL C00595 V=7.0 ACC=20 DEC=20
MOVL C00596 V=7.0 ACC=20 DEC=20
MOVL C00597 V=7.0 ACC=20 DEC=20
MOVL C00598 V=7.0 ACC=20 DEC=20
MOVL C00599 V=7.0 ACC=20 DEC=20
MOVL C00600 V=7.0 ACC=20 DEC=20
MOVL C00601 V=7.0 ACC=20 DEC=20
MOVL C00602 V=7.0 ACC=20 DEC=20
MOVL C00603 V=11.0 ACC=20 DEC=20
MOVC C00604 V=11.0 ACC=20 DEC=20
MOVC C00605 V=11.0 ACC=20 DEC=20
MOVC C00606 V=11.0 ACC=20 DEC=20
MOVL C00607 V=7.0 ACC=20 DEC=20
MOVL C00608 V=7.0 ACC=20 DEC=20
MOVL C00609 V=7.0 ACC=20 DEC=20
MOVL C00610 V=7.0 ACC=20 DEC=20
MOVL C00611 V=7.0 ACC=20 DEC=20
MOVL C00612 V=7.0 ACC=20 DEC=20
MOVL C00613 V=7.0 ACC=20 DEC=20
MOVL C00614 V=7.0 ACC=20 DEC=20
MOVL C00615 V=7.0 ACC=20 DEC=20
MOVL C00616 V=7.0 ACC=20 DEC=20
MOVL C00617 V=7.0 ACC=20 DEC=20
MOVL C00618 V=7.0 ACC=20 DEC=20
MOVL C00619 V=7.0 ACC=20 DEC=20
MOVL C00620 V=7.0 ACC=20 DEC=20
MOVL C00621 V=7.0 ACC=20 DEC=20
MOVL C00622 V=7.0 ACC=20 DEC=20
MOVL C00623 V=7.0 ACC=20 DEC=20
MOVL C00624 V=7.0 ACC=20 DEC=20
MOVL C00625 V=7.0 ACC=20 DEC=20
MOVL C00626 V=7.0 ACC=20 DEC=20
MOVL C00627 V=7.0 ACC=20 DEC=20
MOVL C00628 V=7.0 PL=1
MOVL C00629 V=7.0 ACC=20 DEC=20
MOVL C00630 V=7.0 ACC=20 DEC=20
MOVL C00631 V=7.0 ACC=20 DEC=20
MOVL C00632 V=7.0 ACC=20 DEC=20
MOVL C00633 V=7.0 ACC=20 DEC=20
MOVL C00634 V=7.0 ACC=20 DEC=20
MOVL C00635 V=7.0 ACC=20 DEC=20
MOVL C00636 V=7.0 ACC=20 DEC=20
MOVL C00637 V=7.0 ACC=20 DEC=20
MOVL C00638 V=7.0 ACC=20 DEC=20
ARCOF
TIMER T=30
MOVL C00639 V=11.0 ACC=20 DEC=20
*LAG8
MACRO1 MJ#(0) ARGF2
ARCON
MOVL C00640 V=7.0 ACC=20 DEC=20
MOVL C00641 V=7.0 ACC=20 DEC=20
MOVL C00642 V=7.0 ACC=20 DEC=20
MOVL C00643 V=7.0 ACC=20 DEC=20
MOVL C00644 V=7.0 ACC=20 DEC=20
MOVL C00645 V=7.0 ACC=20 DEC=20
MOVL C00646 V=7.0 ACC=20 DEC=20
MOVL C00647 V=7.0 ACC=20 DEC=20
MOVL C00648 V=7.0 ACC=20 DEC=20
MOVL C00649 V=7.0 PL=1
MOVL C00650 V=7.0 ACC=20 DEC=20
MOVL C00651 V=7.0 ACC=20 DEC=20
MOVL C00652 V=7.0 ACC=20 DEC=20
MOVL C00653 V=7.0 ACC=20 DEC=20
MOVL C00654 V=7.0 ACC=20 DEC=20
MOVL C00655 V=7.0 ACC=20 DEC=20
MOVL C00656 V=7.0 ACC=20 DEC=20
MOVL C00657 V=7.0 ACC=20 DEC=20
MOVL C00658 V=7.0 ACC=20 DEC=20
MOVL C00659 V=7.0 ACC=20 DEC=20
MOVL C00660 V=7.0 ACC=20 DEC=20
MOVL C00661 V=7.0 ACC=20 DEC=20
MOVL C00662 V=7.0 ACC=20 DEC=20
MOVL C00663 V=7.0 ACC=20 DEC=20
MOVL C00664 V=7.0 ACC=20 DEC=20
MOVL C00665 V=7.0 ACC=20 DEC=20
MOVL C00666 V=7.0 ACC=20 DEC=20
MOVL C00667 V=7.0 ACC=20 DEC=20
MOVL C00668 V=7.0 ACC=20 DEC=20
MOVL C00669 V=7.0 ACC=20 DEC=20
MOVL C00670 V=7.0 ACC=20 DEC=20
MOVL C00671 V=11.0 ACC=20 DEC=20
MOVC C00672 V=11.0 ACC=20 DEC=20
MOVC C00673 V=11.0 ACC=20 DEC=20
MOVC C00674 V=11.0 ACC=20 DEC=20
MOVL C00675 V=7.0 ACC=20 DEC=20
MOVL C00676 V=7.0 ACC=20 DEC=20
MOVL C00677 V=7.0 ACC=20 DEC=20
MOVL C00678 V=7.0 ACC=20 DEC=20
MOVL C00679 V=7.0 ACC=20 DEC=20
MOVL C00680 V=7.0 ACC=20 DEC=20
MOVL C00681 V=7.0 ACC=20 DEC=20
MOVL C00682 V=7.0 ACC=20 DEC=20
MOVL C00683 V=7.0 ACC=20 DEC=20
MOVL C00684 V=7.0 ACC=20 DEC=20
MOVL C00685 V=7.0 ACC=20 DEC=20
MOVL C00686 V=7.0 ACC=20 DEC=20
MOVL C00687 V=7.0 ACC=20 DEC=20
MOVL C00688 V=7.0 ACC=20 DEC=20
MOVL C00689 V=7.0 ACC=20 DEC=20
MOVL C00690 V=7.0 ACC=20 DEC=20
MOVL C00691 V=7.0 ACC=20 DEC=20
MOVL C00692 V=7.0 ACC=20 DEC=20
MOVL C00693 V=7.0 ACC=20 DEC=20
MOVL C00694 V=7.0 ACC=20 DEC=20
MOVL C00695 V=7.0 ACC=20 DEC=20
MOVL C00696 V=7.0 PL=1
MOVL C00697 V=7.0 ACC=20 DEC=20
MOVL C00698 V=7.0 ACC=20 DEC=20
MOVL C00699 V=7.0 ACC=20 DEC=20
MOVL C00700 V=7.0 ACC=20 DEC=20
MOVL C00701 V=7.0 ACC=20 DEC=20
MOVL C00702 V=7.0 ACC=20 DEC=20
MOVL C00703 V=7.0 ACC=20 DEC=20
MOVL C00704 V=7.0 ACC=20 DEC=20
MOVL C00705 V=7.0 ACC=20 DEC=20
MOVL C00706 V=11.0 ACC=20 DEC=20
MOVC C00707 V=11.0 ACC=20 DEC=20
MOVC C00708 V=11.0 ACC=20 DEC=20
MOVC C00709 V=11.0 ACC=20 DEC=20
MOVL C00710 V=7.0 ACC=20 DEC=20
MOVL C00711 V=7.0 ACC=20 DEC=20
MOVL C00712 V=7.0 ACC=20 DEC=20
MOVL C00713 V=7.0 ACC=20 DEC=20
MOVL C00714 V=7.0 ACC=20 DEC=20
MOVL C00715 V=7.0 ACC=20 DEC=20
MOVL C00716 V=7.0 ACC=20 DEC=20
MOVL C00717 V=7.0 ACC=20 DEC=20
MOVL C00718 V=7.0 ACC=20 DEC=20
MOVL C00719 V=7.0 ACC=20 DEC=20
MOVL C00720 V=7.0 ACC=20 DEC=20
MOVL C00721 V=7.0 ACC=20 DEC=20
MOVL C00722 V=7.0 ACC=20 DEC=20
MOVL C00723 V=7.0 ACC=20 DEC=20
MOVL C00724 V=7.0 ACC=20 DEC=20
MOVL C00725 V=7.0 ACC=20 DEC=20
MOVL C00726 V=7.0 ACC=20 DEC=20
MOVL C00727 V=7.0 ACC=20 DEC=20
MOVL C00728 V=7.0 ACC=20 DEC=20
MOVL C00729 V=7.0 ACC=20 DEC=20
ARCOF
TIMER T=30
MOVL C00730 V=11.0 ACC=20 DEC=20
*LAG9
MACRO1 MJ#(0) ARGF2
ARCON
MOVL C00731 V=7.0 ACC=20 DEC=20
MOVL C00732 V=7.0 ACC=20 DEC=20
MOVL C00733 V=7.0 ACC=20 DEC=20
MOVL C00734 V=7.0 ACC=20 DEC=20
MOVL C00735 V=7.0 ACC=20 DEC=20
MOVL C00736 V=7.0 ACC=20 DEC=20
MOVL C00737 V=7.0 ACC=20 DEC=20
MOVL C00738 V=7.0 ACC=20 DEC=20
MOVL C00739 V=7.0 ACC=20 DEC=20
MOVL C00740 V=7.0 ACC=20 DEC=20
MOVL C00741 V=7.0 ACC=20 DEC=20
MOVL C00742 V=7.0 ACC=20 DEC=20
MOVL C00743 V=7.0 ACC=20 DEC=20
MOVL C00744 V=7.0 ACC=20 DEC=20
MOVL C00745 V=7.0 ACC=20 DEC=20
MOVL C00746 V=7.0 ACC=20 DEC=20
MOVL C00747 V=7.0 ACC=20 DEC=20
MOVL C00748 V=7.0 ACC=20 DEC=20
MOVL C00749 V=7.0 ACC=20 DEC=20
MOVL C00750 V=11.0 ACC=20 DEC=20
MOVC C00751 V=11.0 ACC=20 DEC=20
MOVC C00752 V=11.0 ACC=20 DEC=20
MOVC C00753 V=11.0 ACC=20 DEC=20
MOVL C00754 V=7.0 ACC=20 DEC=20
MOVL C00755 V=7.0 ACC=20 DEC=20
MOVL C00756 V=7.0 ACC=20 DEC=20
MOVL C00757 V=7.0 ACC=20 DEC=20
MOVL C00758 V=7.0 ACC=20 DEC=20
MOVL C00759 V=7.0 ACC=20 DEC=20
MOVL C00760 V=7.0 ACC=20 DEC=20
MOVL C00761 V=7.0 ACC=20 DEC=20
MOVL C00762 V=7.0 ACC=20 DEC=20
MOVL C00763 V=7.0 PL=1
MOVL C00764 V=7.0 ACC=20 DEC=20
MOVL C00765 V=7.0 ACC=20 DEC=20
MOVL C00766 V=7.0 ACC=20 DEC=20
MOVL C00767 V=7.0 ACC=20 DEC=20
MOVL C00768 V=7.0 ACC=20 DEC=20
MOVL C00769 V=7.0 ACC=20 DEC=20
MOVL C00770 V=7.0 ACC=20 DEC=20
MOVL C00771 V=7.0 ACC=20 DEC=20
MOVL C00772 V=7.0 ACC=20 DEC=20
MOVL C00773 V=7.0 ACC=20 DEC=20
MOVL C00774 V=7.0 ACC=20 DEC=20
MOVL C00775 V=7.0 ACC=20 DEC=20
MOVL C00776 V=7.0 ACC=20 DEC=20
MOVL C00777 V=7.0 ACC=20 DEC=20
MOVL C00778 V=7.0 ACC=20 DEC=20
MOVL C00779 V=7.0 ACC=20 DEC=20
MOVL C00780 V=7.0 ACC=20 DEC=20
MOVL C00781 V=7.0 ACC=20 DEC=20
MOVL C00782 V=7.0 ACC=20 DEC=20
MOVL C00783 V=7.0 ACC=20 DEC=20
MOVL C00784 V=7.0 ACC=20 DEC=20
MOVL C00785 V=11.0 ACC=20 DEC=20
MOVC C00786 V=11.0 ACC=20 DEC=20
MOVC C00787 V=11.0 ACC=20 DEC=20
MOVC C00788 V=11.0 ACC=20 DEC=20
MOVL C00789 V=7.0 ACC=20 DEC=20
MOVL C00790 V=7.0 ACC=20 DEC=20
MOVL C00791 V=7.0 ACC=20 DEC=20
MOVL C00792 V=7.0 ACC=20 DEC=20
MOVL C00793 V=7.0 ACC=20 DEC=20
MOVL C00794 V=7.0 ACC=20 DEC=20
MOVL C00795 V=7.0 ACC=20 DEC=20
MOVL C00796 V=7.0 ACC=20 DEC=20
MOVL C00797 V=7.0 ACC=20 DEC=20
MOVL C00798 V=7.0 ACC=20 DEC=20
MOVL C00799 V=7.0 ACC=20 DEC=20
MOVL C00800 V=7.0 ACC=20 DEC=20
MOVL C00801 V=7.0 ACC=20 DEC=20
MOVL C00802 V=7.0 ACC=20 DEC=20
MOVL C00803 V=7.0 ACC=20 DEC=20
MOVL C00804 V=7.0 ACC=20 DEC=20
MOVL C00805 V=7.0 ACC=20 DEC=20
MOVL C00806 V=7.0 ACC=20 DEC=20
MOVL C00807 V=7.0 ACC=20 DEC=20
MOVL C00808 V=7.0 ACC=20 DEC=20
MOVL C00809 V=7.0 ACC=20 DEC=20
MOVL C00810 V=7.0 PL=1
MOVL C00811 V=7.0 ACC=20 DEC=20
MOVL C00812 V=7.0 ACC=20 DEC=20
MOVL C00813 V=7.0 ACC=20 DEC=20
MOVL C00814 V=7.0 ACC=20 DEC=20
MOVL C00815 V=7.0 ACC=20 DEC=20
MOVL C00816 V=7.0 ACC=20 DEC=20
MOVL C00817 V=7.0 ACC=20 DEC=20
MOVL C00818 V=7.0 ACC=20 DEC=20
MOVL C00819 V=7.0 ACC=20 DEC=20
MOVL C00820 V=7.0 ACC=20 DEC=20
ARCOF
TIMER T=30
MOVL C00821 V=11.0 ACC=20 DEC=20
*LAG10
MACRO1 MJ#(0) ARGF2
ARCON
MOVL C00822 V=7.0 ACC=20 DEC=20
MOVL C00823 V=7.0 ACC=20 DEC=20
MOVL C00824 V=7.0 ACC=20 DEC=20
MOVL C00825 V=7.0 ACC=20 DEC=20
MOVL C00826 V=7.0 ACC=20 DEC=20
MOVL C00827 V=7.0 ACC=20 DEC=20
MOVL C00828 V=7.0 ACC=20 DEC=20
MOVL C00829 V=7.0 ACC=20 DEC=20
MOVL C00830 V=7.0 ACC=20 DEC=20
MOVL C00831 V=7.0 PL=1
MOVL C00832 V=7.0 ACC=20 DEC=20
MOVL C00833 V=7.0 ACC=20 DEC=20
MOVL C00834 V=7.0 ACC=20 DEC=20
MOVL C00835 V=7.0 ACC=20 DEC=20
MOVL C00836 V=7.0 ACC=20 DEC=20
MOVL C00837 V=7.0 ACC=20 DEC=20
MOVL C00838 V=7.0 ACC=20 DEC=20
MOVL C00839 V=7.0 ACC=20 DEC=20
MOVL C00840 V=7.0 ACC=20 DEC=20
MOVL C00841 V=7.0 ACC=20 DEC=20
MOVL C00842 V=7.0 ACC=20 DEC=20
MOVL C00843 V=7.0 ACC=20 DEC=20
MOVL C00844 V=7.0 ACC=20 DEC=20
MOVL C00845 V=7.0 ACC=20 DEC=20
MOVL C00846 V=7.0 ACC=20 DEC=20
MOVL C00847 V=7.0 ACC=20 DEC=20
MOVL C00848 V=7.0 ACC=20 DEC=20
MOVL C00849 V=7.0 ACC=20 DEC=20
MOVL C00850 V=7.0 ACC=20 DEC=20
MOVL C00851 V=7.0 ACC=20 DEC=20
MOVL C00852 V=7.0 ACC=20 DEC=20
MOVL C00853 V=11.0 ACC=20 DEC=20
MOVC C00854 V=11.0 ACC=20 DEC=20
MOVC C00855 V=11.0 ACC=20 DEC=20
MOVC C00856 V=11.0 ACC=20 DEC=20
MOVL C00857 V=7.0 ACC=20 DEC=20
MOVL C00858 V=7.0 ACC=20 DEC=20
MOVL C00859 V=7.0 ACC=20 DEC=20
MOVL C00860 V=7.0 ACC=20 DEC=20
MOVL C00861 V=7.0 ACC=20 DEC=20
MOVL C00862 V=7.0 ACC=20 DEC=20
MOVL C00863 V=7.0 ACC=20 DEC=20
MOVL C00864 V=7.0 ACC=20 DEC=20
MOVL C00865 V=7.0 ACC=20 DEC=20
MOVL C00866 V=7.0 ACC=20 DEC=20
MOVL C00867 V=7.0 ACC=20 DEC=20
